(* IEC 61131-3 sources: daoli-st-library/DL_Motion (part 26) *)

(* ---- FB_DL_WindingTensionCtrl.st ---- *)
(*==============================================================================
 * 组件名称 (Component)  : FB_DL_WindingTensionCtrl
 * 所属子库 (Sublibrary) : DL_Motion
 * 当前版本 (Version)    : 1.0.1
 * 组件分类 (Category)   : 功能块（FUNCTION_BLOCK）· 卷绕工艺族 · 锥度张力闭环
 * 兼容性   (Platform)   : CODESYS 3.5 / TwinCAT 3 / 汇川 InoProShop / Schneider
 *                         Machine Expert；仅依赖 Standard.library（R_TRIG / LIMIT /
 *                         MIN / MAX / ABS / 标准类型转换）
 * 功能描述 (Function)   : 卷绕张力给定合成器。基准张力 = 目标张力 乘 锥度系数（随
 *                         机组直径由 1.0 平滑衰减到 1-K），摆辊位置误差经纯比例
 *                         修正环折算成张力修正量，两层相加后限幅输出，可直接送
 *                         比例阀或伺服转矩限幅入口。卷径可由线速度与角速度反算，
 *                         也可由外部注入。
 * 与既有件边界 (Boundary): FB_DL_WindingTraverse 做排线横动与卷径递推，不含张力
 *                         闭环；FC_DL_CoilDiameterCalc 只做单点几何反算（无状态、
 *                         无记忆）；本件是张力控制层，把二者的能力按需组装。本件
 *                         的相位枚举是工艺相位（闭环 / 开环降级），不是轴状态，轴
 *                         状态机仍归 I_DL_MotionAxis 的 PLCopen 语义，两者严禁合并。
 * 设计要点 (Key notes)  :
 *   ① 降级必须显式：摆辊反馈丢失时进 eOpenLoop 并上报 02D0，只输出锥度基准张力，
 *      不静默沿用上次闭环输出，也不静默把自己当闭环继续算；
 *   ② 修正加在基准上而非串接：摆辊失反馈时仍有锥度张力可用，失反馈不丢张力；
 *   ③ 锥度分母双重校验：满卷直径减卷芯直径小于容差即判退化，系数置 1.0 并上报
 *      01C1，绝不做出除以零的动作；系数再钳到 [1-K, 1.0]，K 自身先钳到 [0, 1]；
 *   ④ 卷径无效沿用上次有效值：转速低于门限时几何反算不可信（编码器低频量化），
 *      沿用上次有效值并累计连续无效次数，超限才升级为 02D1 锁存；
 *   ⑤ 无扰投切：开环恢复闭环时先给 PID 两拍跟踪（跟踪值 0，跟踪窗内过程值同步
 *      取基准以保偏差为零），跟踪结束积分残量为零，比例作用全量恢复；
 *      杜绝投切瞬间张力跳变；
 *   ⑥ 纯比例修正环：PID 实例积分与微分时间均给零，卷径时变工况下不会被积分饱和
 *      拖住。
 * 开源溯源 (Origin)     : 参考 lgf-technology、s7-motion 公开手册与 PLCopen 运动
 *                         控制规范中卷绕张力控制的功能分类与参数域（张力设定、锥度
 *                         系数、摆辊修正、卷径来源四段入口形态），只借分类、参数域
 *                         与命名组织，clean-room 实现，不构成衍生作品。引脚命名、
 *                         枚举、状态跃迁、故障码与合成公式 100% 自有。
 * 依赖     (Depends)    : DL_Algo 已入库件 FB_DL_PidController（拍级 PID，输出域
 *                         经 rOutMin / rOutMax 取 −1~+1 归一化）、
 *                         FC_DL_CoilDiameterCalc（几何反算，入口米制、出口米制，
 *                         本件负责毫米与米换算）。层次合法：Motion 依赖 Algo。
 * 状态迁移 (Transitions):
 *   eIdle      -- bEnable 且 bRun 且摆辊反馈有效 -----------> eClosedLoop（bInControl）
 *   eIdle      -- bEnable 且 bRun 且摆辊反馈无效 -----------> eOpenLoop（02D0 显式降级）
 *   eClosedLoop-- 摆辊反馈丢失 -----------------------------> eOpenLoop（02D0）
 *   eOpenLoop  -- 摆辊反馈连续 3 拍在物理域内 ---------------> eClosedLoop（跟踪投切）
 *   eClosedLoop-- 卷径连续无效次数超限 ---------------------> eFault（02D1 锁存）
 *   eOpenLoop  -- 卷径连续无效次数超限 ---------------------> eFault（02D1 锁存）
 *   任何运行态 -- NOT bEnable 或 NOT bRun ------------------> eIdle（输出 0，PID 复位）
 *   eFault     -- bReset 上升沿 ----------------------------> eIdle
 *   非法枚举值 -- CASE ELSE 兜底 ---------------------------> eFault（复用 02D1）
 * 码位表 (Error codes)  :
 *   16#0004_01C0【信息级】卷径无效（无有效反算或注入非法），已沿用上次有效值；
 *   16#0004_01C1【信息级】锥度系数分母退化或系数超界，已钳位；
 *   16#0004_01C2【信息级】张力输出限幅生效，输出被钳到张力域边界；
 *   16#0004_02D0【故障级】摆辊反馈丢失（非有限值或超机械行程），降级开环；
 *   16#0004_02D1【故障级】卷径连续无效超限（几何法已不可信），锁存待复位。
 *   信息级码只进 uErrorId，不置 bError；02D0 虽为故障级但只降级不停机（bError
 *   置位以提示上游），02D1 进 eFault 锁存。
 * 验收向量 (Acceptance):
 *   V1 锥度：K 0.5、卷芯 200 mm、满卷 1000 mm、实际 800 mm → 系数 0.625；
 *   V2 基准张力：同上且设定 100 N → 基准 62.5 N；
 *   V3 摆辊修正：误差 +2.0 mm、增益 0.5（归一化）、修正满量程 1.0 N → 修正 +1.0 N，
 *      输出 63.5 N；
 *   V4 满卷：实际 1000 mm、设定 100 N → 系数 0.5，基准 50.0 N；
 *   V5 卷径反算：线速 120 米每分、转速 60 转每分、直连 → 卷径约 636.6 mm；
 *   V6 卷径无效：转速 0 → 沿用上次有效卷径，码 01C0，bError 为 FALSE；
 *   V7 反馈丢失：摆辊位置 9999.0 mm → 输出等于基准（不加修正），码 02D0，
 *      bError 为 TRUE，bInControl 为 FALSE。
 * 已知限制 (Limits)     : ① 卷径反算用直连传动比 1.0（机械传动比应由卷径件入口
 *                         承载，本件不重复定义）；② 张力闭环是归一化纯比例修正，
 *                         不做卷径前馈，加减速段的动态偏差仍需现场调 fPidKp；
 *                         ③ 本件不构成安全功能，断带与超张力保护必须由硬件与
 *                         认证安全回路承担。
 * 规格偏离 (Deviation)  : ① 规格伪码把 fPidKp 原样送 PID，同时要求「摆辊正误差得
 *                         正修正」，二者符号相反；本实现送 −ABS(fPidKp)，依托 PID
 *                         件已文档化的「负增益即反作用」特性，令正误差得正修正，
 *                         与验收向量 V3 一致；② 规格成员名 nInvalidDiaCnt 定义类型
 *                         为 UDINT，与「无符号量 u 前缀」红线冲突，改名
 *                         uInvalidDiaCnt（语义不变）；③ 规格未规定故障态张力输出，
 *                         本实现取 0.0 安全值；④ 规格未覆盖「使能瞬间反馈已丢失」
 *                         路径，本实现显式进 eOpenLoop 并带 02D0，不得静默入闭环。
 * 红线自检 (Redline)    : R1 零全局变量表 / 零外部变量声明 / 零物理地址 ✓
 *                         R2 零占位符 ✓ ｜ R3 纯 IEC 61131-3 ✓
 *                         R4 防除零（锥度分母、转速门限）、防越界（卷径钳位）、
 *                         浮点容差（系数域与限幅判定）✓
 *                         R5 声明行 100% 中英双语同行注释 ✓
 *                         R6 ENUM + CASE 且 ELSE 兜底，四态各自有标签 ✓
 *                         R7 R_TRIG 与 PID 实例均在主体无条件刷新 ✓
 * 修订历史 (Revision)   :
 *   2026-11-15  v1.0.0  首版入库（Round 11 · DL_Motion 卷绕张力族开族件）
 *   2026-11-15  v1.0.1  R11 总监终审修复：跟踪拍只置位不递减（bTrack 恒真致修正恒零、
 *                       闭环退化为开环），补 eClosedLoop 逐拍递减；跟踪窗内过程值改取
 *                       基准，消除 PID 反算积分残量（原跟踪结束 fInt 恒等于负比例项，
 *                       V3 修正 +1.0 N 不可达）；02D1 判据由大于改为大于等于，与饱和
 *                       计数上限自洽（原判据在计数封顶时永假，锁存永不触发）
 *   2026-11-15  v1.0.1  R11 director final review fix: the tracking counter now decrements
 *                       every closed-loop scan, the process value follows the reference
 *                       inside the tracking window to keep the back-calculated integral at
 *                       zero, and the 02D1 test uses greater-or-equal against the
 *                       saturating counter so the latch can actually engage
 *============================================================================*)
(*-----------------------------------------------------------------------------
 * 调用示例 (Instance guide)：
 *   // fbTensionPid 与 stStat 均由调用方持有，跨周期传入
 *   fbTension(bEnable := bLineRun, bReset := bFaultReset, bRun := bWinding,
 *             fTensionSet := fTensionRecipe, fDancerPos := fDancerFeedback,
 *             fDancerRef := 0.0, fAxisSpeedRpm := fWinderRpm,
 *             fLineSpeed := fLineSpeedAct, fCoreDia := 200.0,
 *             fDiaMax := 1000.0, bUseInjectedDia := FALSE,
 *             fTaperK := 0.50, fPidKp := 0.5, fTrimSpan := 5.0,
 *             fTensionMin := 0.0, fTensionMax := 300.0);
 *   fValveCmd := fbTension.fTensionOut;
 *   注：fbTensionPid 只允许本块调用，外部不要再对该实例赋值引脚，否则归一化
 *       输出域会被覆盖，修正量会放大一百倍。
 *----------------------------------------------------------------------------*)
(*-----------------------------------------------------------------------------
 * 常见误用与现场提示 (Field notes)：
 *   1 fTaperK 给 0 表示无锥度（全程恒张力），给 1 表示满卷张力降到零，后者在
 *     实际工艺中通常不可用，建议上限取 0.7。
 *   2 摆辊反馈量程必须与 fDancerRef 同一基准：本块用绝对值 500 mm 判机械不可能
 *     值，若机械行程超过 500 mm，请把 DL_DANCER_LIMIT 调大后重新入库。
 *   3 卷径连续无效 50 次即锁存 02D1：停机不转时卷径无效属正常（信息级 01C0），
 *     只要 bRun 撤除就不会累计，现场不要把停机误判为故障。
 *   4 开环降级期间张力只随卷径变化，摆辊会漂到机械限位，现场必须给摆辊限位
 *     开关并把其信号接入上位联锁，本块不做摆辊位置保护。
 *   5 张力上下限写反时本块自动对调，但不会报警，调试期请核对 fTensionMin 与
 *     fTensionMax 的实际取值。
 *----------------------------------------------------------------------------*)
(*-----------------------------------------------------------------------------
 * 枚举: E_DL_TensionPhase（归属 DL_Motion，与本功能块同文件发布）
 * 含义: 张力工艺相位。eOpenLoop 是显式降级态而非故障态，二者不可混用。
 *----------------------------------------------------------------------------*)
{attribute 'strict'}
{attribute 'qualified_only'}
TYPE E_DL_TensionPhase :
(
    eIdle       := 0,   // 空闲：未使能或未运行，张力输出 0，PID 复位 / Idle: disabled or not running, tension output zero, PID reset
    eOpenLoop   := 10,  // 开环降级：摆辊反馈不可用，只出锥度基准张力 / Open loop degraded: dancer feedback unusable, taper base only
    eClosedLoop := 20,  // 闭环运行：基准张力加摆辊比例修正 / Closed loop: base tension plus dancer proportional trim
    eFault      := 99   // 故障锁存：卷径几何法不可信，仅复位沿退出 / Fault latched: diameter geometry untrusted, exits on reset edge only
) UINT;
END_TYPE
(*-----------------------------------------------------------------------------
 * 结构体: ST_DL_WindingStat（归属 DL_Motion，与本功能块同文件发布）
 * 含义: 卷绕统计，由调用方持有并可持久化到配方域。
 *----------------------------------------------------------------------------*)
TYPE ST_DL_WindingStat :
STRUCT
    fTensionAvg     : REAL;   // 张力滑动均值 [N]，一阶指数平均，仅闭环期更新 / Tension running average in newtons, updated in closed loop only
    uInvalidDiaCnt  : UDINT;  // 卷径连续无效次数 [次]，任一有效反算即清零 / Consecutive invalid diameter count, cleared by any valid result
    tRunTime        : TIME;   // 闭环累计运行时长 [ms]，按任务周期累加 / Accumulated closed-loop runtime in milliseconds
END_STRUCT
END_TYPE

(*==============================================================================
 * 功能块: FB_DL_WindingTensionCtrl
 * 调用约定: 每扫描周期无条件调用一次；PID 实例在主体末尾无条件调用。
 * 无状态泄漏: 状态驻留实例私有 VAR 与调用方持有的 stStat / fbTensionPid。
 *============================================================================*)
FUNCTION_BLOCK FB_DL_WindingTensionCtrl
VAR_INPUT
    bEnable          : BOOL := FALSE;        // 总使能 [BOOL]，FALSE 时输出 0 并复位 PID / Master enable, FALSE zeroes the output and resets the PID
    bReset           : BOOL := FALSE;        // 复位 [BOOL]，上升沿复位故障、计数与 PID / Reset, rising edge clears fault, counters and the PID
    bRun             : BOOL := FALSE;        // 卷绕运行中 [BOOL]，FALSE 时张力给定保持 0 / Winding running flag, FALSE holds the tension command at zero
    fTensionSet      : REAL := 0.0;          // 目标张力（满卷前基准）[N]，域 0.0~500.0 / Base tension setpoint in newtons, range zero to five hundred
    fDancerPos       : REAL := 0.0;          // 摆辊实际位置 [mm]，0 为机械中位，绝对值超 500 判失效 / Dancer actual position in millimetres, zero at mechanical centre
    fDancerRef       : REAL := 0.0;          // 摆辊中位基准 [mm]，非有限值按 0 处理 / Dancer centre reference in millimetres, non-finite treated as zero
    fAxisSpeedRpm    : REAL := 0.0;          // 卷轴转速 [转每分]，低于 1.0 视为不可反算 / Winder shaft speed in revolutions per minute, below one is untrusted
    fLineSpeed       : REAL := 0.0;          // 线速度 [米每分]，与卷径件入口同单位 / Line speed in metres per minute, same unit as the diameter function input
    fCoreDia         : REAL := 200.0;        // 卷芯直径 [mm]，域 10.0~3000.0 / Core diameter in millimetres, range ten to three thousand
    fDiaMax          : REAL := 1000.0;       // 满卷直径 [mm]，必须大于卷芯直径，否则锥度退化 / Full roll diameter in millimetres, must exceed the core diameter
    fDiaInjected     : REAL := 0.0;          // 外部注入卷径 [mm]，视觉或上位机来源 / Injected diameter in millimetres from vision or a host system
    bUseInjectedDia  : BOOL := FALSE;        // 卷径来源选择 [BOOL]，TRUE 用注入值，FALSE 由速度比反算 / Diameter source, TRUE uses the injected value
    fThickness       : REAL := 0.10;         // 材料厚度 [mm]，供卷径件层数积分 / Material thickness in millimetres, used by the layer integral
    fTaperK          : REAL := 0.50;         // 锥度系数 [无量纲 0~1]，满卷张力降至 1-K 倍 / Taper coefficient, full roll tension falls to one minus K
    fPidKp           : REAL := 0.5;          // 摆辊修正归一化增益 [每毫米]，输出域 −1~+1，取绝对值后反作用 / Normalised dancer gain per millimetre, absolute value used with reverse action
    fTrimSpan        : REAL := 1.0;          // 修正满量程 [N]，归一化输出乘该值即张力修正 / Trim span in newtons, the normalised output multiplied by this value
    fTensionMin      : REAL := 0.0;          // 张力输出下限 [N]，与上限对调时自动修复 / Tension lower limit in newtons, swapped limits are repaired
    fTensionMax      : REAL := 500.0;        // 张力输出上限 [N]，等于下限时输出被钉死 / Tension upper limit in newtons, an equal limit pins the output
END_VAR
VAR_OUTPUT
    fTensionOut      : REAL := 0.0;          // 张力给定输出 [N]，送比例阀或转矩限幅入口 / Tension command output in newtons for a proportional valve or torque limit
    fDiaAct          : REAL := 0.0;          // 当前生效卷径 [mm]，已钳入物理域 / Effective diameter in millimetres, clamped into the physical range
    fTaperFactor     : REAL := 1.0;          // 实际锥度系数 [无量纲]，域 1-K~1.0 / Effective taper factor, range one minus K to one
    fDancerErr       : REAL := 0.0;          // 摆辊位置误差 [mm]，等于实测减基准 / Dancer position error in millimetres, measured minus reference
    eState           : E_DL_TensionPhase := E_DL_TensionPhase.eIdle; // 主状态机当前态 [枚举] / Current state of the main state machine
    bInControl       : BOOL := FALSE;        // 张力闭环生效 [BOOL]，仅 eClosedLoop 为 TRUE / Closed-loop tension active, TRUE only in the closed-loop state
    bError           : BOOL := FALSE;        // 故障标志 [BOOL]，故障级码或降级态置位，信息级码不置位 / Fault flag, set by fault-level codes or the degraded state
    uErrorId         : UDINT := 0;           // 事件或故障码 [段位 0004_01Cx 与 0004_02Dx]，0 表示无事件 / Event or fault code in the 0004 bands, zero means none
    fDiaLastValid    : REAL := 0.0;          // 最近一次有效卷径 [mm]，0 表示尚无有效值 / Last valid diameter in millimetres, zero means none yet
END_VAR
VAR_IN_OUT
    fbTensionPid     : FB_DL_PidController;  // 摆辊修正环 PID 实例 [FB]，由调用方持有且只允许本块调用 / Dancer trim PID instance held by the caller and driven only by this block
    stStat           : ST_DL_WindingStat;    // 跨周期卷绕统计 [结构体]，由调用方持有 / Persistent winding statistics held by the caller
END_VAR
VAR
    bInit            : BOOL := FALSE;        // 首扫完成标志 [BOOL]，初值 FALSE，判据恒为 NOT bInit / First-scan done flag, initial FALSE, judged by NOT bInit
    bDancerOk        : BOOL := FALSE;        // 摆辊反馈有效判据 [BOOL]，逐拍重算 / Dancer feedback verdict, recomputed every scan
    bDancerLost      : BOOL := FALSE;        // 摆辊反馈丢失标志 [BOOL]，降级原因量 / Dancer feedback lost flag, the explicit degradation reason
    bAvgInit         : BOOL := FALSE;        // 张力均值首样本标志 [BOOL]，避免从 0 起算 / Tension average first-sample flag, avoids averaging from zero
    nRecoverCnt      : INT := 0;             // 反馈恢复连续拍计数 [拍]，满 3 拍回闭环 / Consecutive good-feedback counter, three scans restore closed loop
    nTrackSync       : INT := 0;             // 投切跟踪剩余拍数 [拍]，大于 0 时 PID 跟踪 / Remaining tracking scans, the PID tracks while above zero
    fDancerPosEff    : REAL := 0.0;          // 喂给 PID 的摆辊位置 [mm]，失效时以基准值替代 / Dancer position fed to the PID, replaced by the reference when invalid
    fDancerRefEff    : REAL := 0.0;          // 生效摆辊基准 [mm]，已做非有限值防御 / Effective dancer reference after the non-finite defence
    fPidPvEff        : REAL := 0.0;          // 喂给 PID 的过程值 [mm]，跟踪窗口内以基准替代 / Process value fed to the PID, replaced by the reference inside the tracking window
    fTensionSetEff   : REAL := 0.0;          // 生效目标张力 [N]，已做非有限值防御 / Effective tension setpoint after the non-finite defence
    fTrimSpanEff     : REAL := 1.0;          // 生效修正满量程 [N]，取绝对值 / Effective trim span in newtons, absolute value used
    fPidKpEff        : REAL := 0.0;          // 送入 PID 的增益 [每毫米]，取负值实现反作用 / Gain passed to the PID, negated for reverse action
    fCoreDiaEff      : REAL := 200.0;        // 生效卷芯直径 [mm]，钳入物理域 / Effective core diameter in millimetres, clamped into the physical range
    fDiaMaxEff       : REAL := 1000.0;       // 生效满卷直径 [mm]，钳入物理域 / Effective full-roll diameter in millimetres, clamped into the physical range
    fTaperKEff       : REAL := 0.50;         // 生效锥度系数 [无量纲 0~1]，越界钳位 / Effective taper coefficient, clamped into zero to one
    fTaperLow        : REAL := 0.50;         // 锥度系数下限 [无量纲]，等于 1 减生效锥度 / Taper factor lower bound, equal to one minus the effective coefficient
    fTaperRaw        : REAL := 1.0;          // 未钳位的锥度系数 [无量纲]，用于超界判定 / Unclamped taper factor used for the out-of-range test
    fDiaCalc         : REAL := 0.0;          // 卷径反算结果 [mm]，已做米转毫米 / Diameter result in millimetres after the metre conversion
    fDiaLReal        : LREAL := 0.0;         // 卷径件出口绑定值 [米]，LREAL 精度承接 / Diameter bound from the function output in metres at LREAL precision
    fDiaRet          : LREAL := 0.0;         // 卷径件返回值 [米]，函数返回即滤波后卷径 / Diameter function return value in metres, the filtered diameter
    fBase            : REAL := 0.0;          // 锥度基准张力 [N]，等于设定乘锥度系数 / Taper base tension in newtons, setpoint times the taper factor
    fTrim            : REAL := 0.0;          // 摆辊张力修正 [N]，闭环时等于归一化输出乘满量程 / Dancer trim in newtons, the normalised output times the span
    fRawCmd          : REAL := 0.0;           // 未限幅的张力指令 [N]，限幅前中间量 / Unlimited tension command in newtons before clamping
    fLimLow          : REAL := 0.0;          // 生效张力下限 [N]，已做上下对调修复 / Effective tension lower limit after repair
    fLimHigh         : REAL := 500.0;        // 生效张力上限 [N]，已做上下对调修复 / Effective tension upper limit after repair
    fAvgAlpha        : REAL := 0.0;          // 张力均值一阶权重 [无量纲]，由任务周期与时间常数算出 / First-order weight of the tension average
    uErrInfo         : UDINT := 0;           // 本拍瞬时信息码 [段位 0004_01C0~01C2]，逐拍重算 / Transient info code recomputed every scan
    uErrFault        : UDINT := 0;           // 锁存故障码 [段位 0004_02D1]，仅复位清除 / Latched fault code, cleared by reset only
    fbTrigReset      : R_TRIG;               // 复位上升沿检测实例 / Rising edge detector for the reset flag
    fbTrigRun        : R_TRIG;               // 运行上升沿检测实例 / Rising edge detector for the running flag
END_VAR
VAR CONSTANT
    DL_FLOAT_EPS     : REAL := 1.0E-6;       // 浮点判等与判零容差 [无量纲，按比较量量纲同值使用] / Float equality and zero tolerance
    DL_INF_MAX       : REAL := 1.0E30;       // 有限值幅值上限 [无量纲，按各量量纲同值使用] / Finite magnitude upper bound
    DL_RPM_MIN       : REAL := 1.0;          // 卷径反算最小转速 [转每分]，低于此值不反算 / Minimum speed for the inverse diameter calculation
    DL_DIA_MIN       : REAL := 10.0;         // 卷径物理下限 [mm] / Diameter physical lower bound in millimetres
    DL_DIA_MAX       : REAL := 3000.0;       // 卷径物理上限 [mm] / Diameter physical upper bound in millimetres
    DL_DANCER_LIMIT  : REAL := 500.0;        // 摆辊机械行程上限 [mm]，绝对值超此判失效 / Dancer mechanical travel bound in millimetres
    DL_TASK_CYCLE    : REAL := 0.010;        // 主任务周期 [s]，供卷径件变化率换算 / Main task cycle in seconds for the diameter rate
    DL_TASK_TIME     : TIME := T#10MS;       // 主任务周期时间量 [ms]，供运行时长累加 / Main task cycle as a time value for runtime accumulation
    DL_FILTER_TAU    : REAL := 0.50;         // 卷径一阶低通时间常数 [s] / Diameter low-pass time constant in seconds
    DL_INVALID_MAX   : UDINT := 50;          // 卷径连续无效次数上限 [次]，超限锁存 02D1 / Consecutive invalid diameter limit before latching
    DL_RECOVER_N     : INT := 3;             // 反馈恢复确认拍数 [拍]，连续满足才回闭环 / Consecutive good scans required to restore the closed loop
    DL_AVG_TAU       : REAL := 1.0;          // 张力均值时间常数 [s]，一阶平均用 / Tension average time constant in seconds
END_VAR
(*------------------------------------------------------------------------------
 * 段 1｜边沿实例无条件周期刷新（红线 R7：严禁置于 IF 或 CASE 分支内）｜Unconditional edge refresh, never placed inside IF or CASE branches
 *-----------------------------------------------------------------------------*)
fbTrigReset(CLK := bReset);
fbTrigRun(CLK := bRun);
(*------------------------------------------------------------------------------
 * 段 2｜瞬时输出与瞬时码预清零（出口只置位，跨拍残留一律在入口清）｜Pre-clear transient outputs and info codes at scan entry
 *-----------------------------------------------------------------------------*)
bInControl := FALSE;                        // 闭环生效标志预清零 [BOOL] / Pre-clear the closed-loop flag
fTrim      := 0.0;                          // 修正量预清零，开环与空闲不得继承上次值 [N] / Pre-clear the trim so open loop never inherits it
uErrInfo   := 0;                            // 瞬时信息码预清零 [码] / Pre-clear the transient info code
(*------------------------------------------------------------------------------
 * 段 3｜参数域修复（引脚可在线改，故逐拍重算；域非法只钳位不锁存）｜Parameter domain repair, clamping only without latching
 *-----------------------------------------------------------------------------*)
IF fTensionMax < fTensionMin THEN
    fLimLow  := fTensionMax;                // 张力域上下对调修复：下限取原上限 [N] / Repaired lower limit takes the original upper
    fLimHigh := fTensionMin;                // 张力域上下对调修复：上限取原下限 [N] / Repaired upper limit takes the original lower
ELSE
    fLimLow  := fTensionMin;                // 合法下限直通 [N] / Valid lower limit passed through
    fLimHigh := fTensionMax;                // 合法上限直通 [N] / Valid upper limit passed through
END_IF

IF (fTensionSet <> fTensionSet) OR (ABS(fTensionSet) > DL_INF_MAX) THEN
    fTensionSetEff := 0.0;                  // 目标张力非有限 → 0，宁可失张力也不给非法值 [N] / Non-finite setpoint falls back to zero
ELSE
    fTensionSetEff := fTensionSet;          // 合法目标张力直通 [N] / Valid setpoint passed through
END_IF

IF (fTrimSpan <> fTrimSpan) OR (ABS(fTrimSpan) > DL_INF_MAX) THEN
    fTrimSpanEff := 0.0;                    // 修正满量程非有限 → 0，等效关闭摆辊修正 [N] / Non-finite trim span disables the dancer trim
ELSE
    fTrimSpanEff := ABS(fTrimSpan);         // 修正满量程取绝对值 [N] / Absolute trim span
END_IF
// 送入 PID 的增益取负实现反作用：摆辊正误差（上偏）对应增张力，与验收向量 V3 一致
IF (fPidKp <> fPidKp) OR (ABS(fPidKp) > DL_INF_MAX) THEN
    fPidKpEff := 0.0;                       // 增益非有限 → 0，等效关闭修正 [每毫米] / Non-finite gain disables the trim
ELSE
    fPidKpEff := -ABS(fPidKp);              // 取绝对值后取负，负增益即 PID 件的反作用语义 [每毫米] / Absolute value negated for reverse action
END_IF

IF (fDancerRef <> fDancerRef) OR (ABS(fDancerRef) > DL_DANCER_LIMIT) THEN
    fDancerRefEff := 0.0;                   // 摆辊基准非法 → 回机械中位 0 [mm] / Illegal reference falls back to the mechanical centre
ELSE
    fDancerRefEff := fDancerRef;            // 合法基准直通 [mm] / Valid reference passed through
END_IF

IF (fCoreDia <> fCoreDia) OR (ABS(fCoreDia) > DL_INF_MAX) THEN
    fCoreDiaEff := DL_DIA_MIN;              // 卷芯直径非法 → 回物理下限 [mm] / Illegal core diameter falls back to the physical lower bound
ELSE
    fCoreDiaEff := LIMIT(DL_DIA_MIN, fCoreDia, DL_DIA_MAX); // 卷芯直径钳入物理域 [mm] / Core diameter clamped into the physical range
END_IF

IF (fDiaMax <> fDiaMax) OR (ABS(fDiaMax) > DL_INF_MAX) THEN
    fDiaMaxEff := DL_DIA_MAX;               // 满卷直径非法 → 回物理上限 [mm] / Illegal full-roll diameter falls back to the physical upper bound
ELSE
    fDiaMaxEff := LIMIT(DL_DIA_MIN, fDiaMax, DL_DIA_MAX);   // 满卷直径钳入物理域 [mm] / Full-roll diameter clamped into the physical range
END_IF
// 锥度系数域校验：非有限或越出 0~1 一律钳位并置信息级 01C1，绝不带非法系数进公式
IF (fTaperK <> fTaperK) OR (ABS(fTaperK) > DL_INF_MAX) THEN
    fTaperKEff := 0.0;                      // 非有限系数按无锥度处理，先判非数再钳位，避免 NaN 穿过 LIMIT [无量纲] / Non-finite coefficient treated as no taper
    IF bEnable AND bRun THEN
        uErrInfo := 16#0004_01C1;           // 【信息级】锥度系数非有限已按无锥度处理 / Info: non-finite taper coefficient replaced
    END_IF
ELSIF (fTaperK < 0.0) OR (fTaperK > 1.0) THEN
    fTaperKEff := LIMIT(0.0, fTaperK, 1.0); // 越界钳到 0~1 双向钳位 [无量纲] / Two-sided clamp into zero to one
    IF bEnable AND bRun THEN
        uErrInfo := 16#0004_01C1;           // 【信息级】锥度系数超界已钳位 / Info: taper coefficient clamped
    END_IF
ELSE
    fTaperKEff := fTaperK;                  // 合法锥度系数直通 [无量纲] / Valid taper coefficient passed through
END_IF
// 张力均值一阶权重：由任务周期与时间常数算出，分母恒正（时间常数有下限保证）
fAvgAlpha := DL_TASK_CYCLE / (DL_AVG_TAU + DL_TASK_CYCLE); // 均值权重 [无量纲] / First-order average weight
(*------------------------------------------------------------------------------
 * 段 4｜首扫装载（R19 唯一合法范式：bInit 初值 FALSE，判据 NOT bInit）｜First-scan load, the only accepted initialisation pattern
 *-----------------------------------------------------------------------------*)
IF NOT bInit THEN
    stStat.fTensionAvg    := 0.0;           // 张力均值清零，等首个闭环样本直取 [N] / Clear the tension average until the first closed-loop sample
    stStat.uInvalidDiaCnt := 0;             // 卷径无效计数清零 [次] / Clear the invalid diameter counter
    stStat.tRunTime       := T#0S;          // 运行时长清零 [ms] / Clear the accumulated runtime
    fDiaLastValid         := 0.0;           // 有效卷径历史清零，0 表示尚无有效值 [mm] / Clear the valid diameter history
    bDancerLost           := FALSE;         // 反馈丢失标志清零 [BOOL] / Clear the feedback lost flag
    nRecoverCnt           := 0;             // 恢复计数清零 [拍] / Clear the recovery counter
    nTrackSync            := 0;             // 投切跟踪计数清零 [拍] / Clear the tracking counter
    bAvgInit              := FALSE;         // 均值首样本标志清零 [BOOL] / Clear the average first-sample flag
    bInit                 := TRUE;          // 首扫完成置位 [BOOL] / First scan completed
END_IF
(*------------------------------------------------------------------------------
 * 段 5｜复位（清故障、计数与降级标志；PID 由复位引脚同步清除；参数域不动）｜Reset clears the latched fault, counters and degradation flags
 *-----------------------------------------------------------------------------*)
IF fbTrigReset.Q THEN
    uErrFault             := 0;             // 锁存故障码清零 [码] / Clear the latched fault code
    uErrInfo              := 0;             // 瞬时信息码清零 [码] / Clear the transient info code
    stStat.uInvalidDiaCnt := 0;             // 卷径无效计数清零，允许重新起步 [次] / Clear the invalid diameter counter so production can restart
    bDancerLost           := FALSE;         // 反馈丢失标志清零 [BOOL] / Clear the feedback lost flag
    nRecoverCnt           := 0;             // 恢复计数清零 [拍] / Clear the recovery counter
    nTrackSync            := 0;             // 跟踪计数清零 [拍] / Clear the tracking counter
    eState                := E_DL_TensionPhase.eIdle; // 回空闲，等待使能与运行条件 [枚举] / Back to idle waiting for enable and run
END_IF

IF fbTrigRun.Q THEN
    bAvgInit := FALSE;                      // 新一次卷绕启动：张力均值重新直取首样本，不继承上一卷 [BOOL] / New run restarts the tension average instead of inheriting the last roll
END_IF
(*------------------------------------------------------------------------------
 * 段 6｜摆辊反馈有效性判定（非有限值或超机械行程即判失效，显式标记原因）｜Dancer feedback verdict with an explicit reason flag
 *-----------------------------------------------------------------------------*)
bDancerOk := NOT ((fDancerPos <> fDancerPos) OR (ABS(fDancerPos) > DL_DANCER_LIMIT));
IF bDancerOk THEN
    fDancerPosEff := fDancerPos;            // 有效反馈直通，喂给 PID [mm] / Valid feedback passed through to the PID
ELSE
    fDancerPosEff := fDancerRefEff;         // 失效反馈以基准替代，令 PID 偏差为零且 NaN 不扩散 [mm] / Substitute the reference so the PID error stays zero
END_IF
fDancerErr := fDancerPosEff - fDancerRefEff; // 摆辊位置误差，实测减基准 [mm] / Dancer position error, measured minus reference
(*------------------------------------------------------------------------------
 * 段 7｜卷径获取（注入优先；否则按速度比反算；无效沿用上次有效值并计数）｜Diameter acquisition with reuse-on-invalid and consecutive counting
 *-----------------------------------------------------------------------------*)
IF bEnable AND bRun THEN
    IF bUseInjectedDia THEN
        IF (fDiaInjected <> fDiaInjected) OR (ABS(fDiaInjected) > DL_INF_MAX) THEN
            IF fDiaLastValid > DL_FLOAT_EPS THEN
                fDiaAct := fDiaLastValid;   // 注入值非法 → 沿用上次有效卷径 [mm] / Illegal injection reuses the last valid diameter
            ELSE
                fDiaAct := fCoreDiaEff;     // 无历史有效值 → 以卷芯直径兜底，杜绝零卷径除零 [mm] / Fall back to the core diameter when no history exists
            END_IF
            IF stStat.uInvalidDiaCnt < DL_INVALID_MAX THEN
                stStat.uInvalidDiaCnt := stStat.uInvalidDiaCnt + 1; // 连续无效计数累加，封顶后靠 02D1 锁存 [次] / Saturating invalid counter
            END_IF
            uErrInfo := 16#0004_01C0;       // 【信息级】卷径无效已沿用上次有效值 / Info: invalid diameter, last valid value reused
        ELSE
            fDiaAct := LIMIT(DL_DIA_MIN, fDiaInjected, DL_DIA_MAX); // 注入卷径钳入物理域 [mm] / Injected diameter clamped into the physical range
            IF (fDiaInjected < DL_DIA_MIN) OR (fDiaInjected > DL_DIA_MAX) THEN
                uErrInfo := 16#0004_01C0;   // 【信息级】注入卷径超物理域已钳位 / Info: injected diameter clamped
            END_IF
            fDiaLastValid         := fDiaAct; // 记录有效卷径 [mm] / Record the valid diameter
            stStat.uInvalidDiaCnt := 0;     // 有效值出现即清零连续无效计数 [次] / Reset the consecutive counter on any valid value
        END_IF
    ELSE
        IF (fAxisSpeedRpm <> fAxisSpeedRpm) OR (ABS(fAxisSpeedRpm) > DL_INF_MAX)
           OR (fAxisSpeedRpm < DL_RPM_MIN)
           OR (fLineSpeed <> fLineSpeed) OR (ABS(fLineSpeed) > DL_INF_MAX) THEN
            IF fDiaLastValid > DL_FLOAT_EPS THEN
                fDiaAct := fDiaLastValid;   // 低速或入参非法 → 沿用上次有效卷径 [mm] / Low speed or illegal input reuses the last valid diameter
            ELSE
                fDiaAct := fCoreDiaEff;     // 无历史有效值 → 以卷芯直径兜底 [mm] / Fall back to the core diameter
            END_IF
            IF stStat.uInvalidDiaCnt < DL_INVALID_MAX THEN
                stStat.uInvalidDiaCnt := stStat.uInvalidDiaCnt + 1; // 连续无效计数累加 [次] / Saturating invalid counter
            END_IF
            uErrInfo := 16#0004_01C0;       // 【信息级】卷径无效已沿用上次有效值 / Info: invalid diameter, last valid value reused
        ELSE
            // 按已入库卷径件的真实契约调用：入口为米制与秒制，出口绑定滤波后卷径（米）
            fDiaRet := FC_DL_CoilDiameterCalc(
                fLineSpeed := REAL_TO_LREAL(fLineSpeed),              // 米每分，与本件引脚同单位 / Metres per minute, same unit as this pin
                fShaftRpm  := REAL_TO_LREAL(fAxisSpeedRpm),           // 转每分，与卷轴转速同单位 / Revolutions per minute
                fGearRatio := 1.0,                                    // 直连，机械传动比由卷径件入口承载 / Direct drive, the gear ratio belongs to the function input
                fCoreDia   := REAL_TO_LREAL(fCoreDiaEff) / 1000.0,     // 毫米转米 / Millimetres converted to metres
                fThickness := REAL_TO_LREAL(fThickness) / 1000.0,     // 毫米转米 / Millimetres converted to metres
                fPrevDia   := REAL_TO_LREAL(fDiaLastValid) / 1000.0,  // 毫米转米，0 表示无历史 / Millimetres converted to metres, zero means no history
                fTaskCycle := REAL_TO_LREAL(DL_TASK_CYCLE),           // 任务周期，秒 / Task cycle in seconds
                bFilterEn  := TRUE,                                   // 卷径低通使能 / Diameter low-pass enabled
                fFilterTau := REAL_TO_LREAL(DL_FILTER_TAU),           // 低通时间常数，秒 / Low-pass time constant in seconds
                fDia       => fDiaLReal );                            // 出口绑定：滤波后卷径，米 / Bound output, filtered diameter in metres
            fDiaCalc := LREAL_TO_REAL(fDiaLReal * 1000.0);            // 米转毫米，显式转换，出口绑定优先 / Metres converted to millimetres, the bound output is preferred
            IF (fDiaLReal <> fDiaLReal) AND (fDiaRet = fDiaRet) THEN
                fDiaCalc := LREAL_TO_REAL(fDiaRet * 1000.0);          // 绑定值非法而返回值有效 → 退回返回值，兼容平台绑定差异 / Bound value illegal, fall back to the function return
            END_IF
            IF (fDiaCalc <> fDiaCalc) OR (fDiaCalc <= DL_FLOAT_EPS) THEN
                IF fDiaLastValid > DL_FLOAT_EPS THEN
                    fDiaAct := fDiaLastValid; // 反算结果不可用 → 沿用上次有效卷径 [mm] / Unusable result reuses the last valid diameter
                ELSE
                    fDiaAct := fCoreDiaEff;   // 无历史有效值 → 以卷芯直径兜底 [mm] / Fall back to the core diameter
                END_IF
                IF stStat.uInvalidDiaCnt < DL_INVALID_MAX THEN
                    stStat.uInvalidDiaCnt := stStat.uInvalidDiaCnt + 1; // 连续无效计数累加 [次] / Saturating invalid counter
                END_IF
                uErrInfo := 16#0004_01C0;   // 【信息级】反算结果不可用已沿用上次有效值 / Info: unusable result, last valid value reused
            ELSE
                fDiaAct := LIMIT(DL_DIA_MIN, fDiaCalc, DL_DIA_MAX); // 反算卷径钳入物理域 [mm] / Computed diameter clamped into the physical range
                fDiaLastValid         := fDiaAct; // 记录有效卷径 [mm] / Record the valid diameter
                stStat.uInvalidDiaCnt := 0;       // 有效反算即清零连续无效计数 [次] / Reset the consecutive counter on a valid result
            END_IF
        END_IF
    END_IF
ELSE
    IF fDiaLastValid > DL_FLOAT_EPS THEN
        fDiaAct := fDiaLastValid;           // 非运行态不反算，沿用上次有效卷径 [mm] / Not running, reuse the last valid diameter
    ELSE
        fDiaAct := fCoreDiaEff;             // 非运行且无历史 → 以卷芯直径兜底 [mm] / Not running without history falls back to the core diameter
    END_IF
END_IF

// 卷径输出钳位兜底：任何路径都不得把非法值送出（防御性二次确认）
IF (fDiaAct <> fDiaAct) OR (fDiaAct < DL_DIA_MIN) OR (fDiaAct > DL_DIA_MAX) THEN
    fDiaAct := LIMIT(DL_DIA_MIN, fDiaAct, DL_DIA_MAX); // 卷径域二次钳位 [mm] / Second-stage diameter clamp
    IF fDiaAct <> fDiaAct THEN
        fDiaAct := fCoreDiaEff;             // 仍为非法值 → 回卷芯直径 [mm] / Still illegal, fall back to the core diameter
    END_IF
END_IF
(*------------------------------------------------------------------------------
 * 段 8｜锥度系数（分母双重校验，系数双向钳位，退化或超界置 01C1）｜Taper factor with denominator guard and two-sided clamping
 *-----------------------------------------------------------------------------*)
IF ABS(fDiaMaxEff - fCoreDiaEff) <= DL_FLOAT_EPS THEN
    fTaperFactor := 1.0;                    // 满卷等于卷芯：锥度退化，系数取 1.0 防除零 [无量纲] / Degenerate span, unity factor avoids division by zero
    IF bEnable AND bRun THEN
        uErrInfo := 16#0004_01C1;           // 【信息级】锥度分母退化已改置 1.0 / Info: degenerate taper span replaced by unity
    END_IF
ELSE
    fTaperLow := 1.0 - fTaperKEff;          // 锥度系数下限，等于 1 减锥度 [无量纲] / Taper factor lower bound
    fTaperRaw := 1.0 - fTaperKEff * (fDiaAct - fCoreDiaEff) / (fDiaMaxEff - fCoreDiaEff); // 原始锥度系数 [无量纲] / Raw taper factor
    IF (fTaperRaw > 1.0 + DL_FLOAT_EPS) OR (fTaperRaw < fTaperLow - DL_FLOAT_EPS) THEN
        fTaperFactor := LIMIT(fTaperLow, fTaperRaw, 1.0); // 超界钳到 [1-K, 1] [无量纲] / Clamp into the lower bound and one
        IF bEnable AND bRun THEN
            uErrInfo := 16#0004_01C1;       // 【信息级】锥度系数超界已钳位 / Info: taper factor clamped
        END_IF
    ELSE
        fTaperFactor := fTaperRaw;          // 未超界直通 [无量纲] / Raw factor passed through
    END_IF
END_IF
(*------------------------------------------------------------------------------
 * 段 9｜锥度基准张力（修正项后续加在基准上，失反馈也不丢张力）｜Taper base tension, the trim is added on top later
 *-----------------------------------------------------------------------------*)
fBase := fTensionSetEff * fTaperFactor;     // 基准张力＝目标张力乘锥度系数 [N] / Base tension equals setpoint times taper factor
(*------------------------------------------------------------------------------
 * 段 10｜主状态机（红线 R6：ENUM + CASE + ELSE 兜底，四态各有标签）｜Main state machine with mandatory ELSE fallback and four labelled states
 *-----------------------------------------------------------------------------*)
CASE eState OF

    E_DL_TensionPhase.eIdle:                // 空闲：等使能与运行条件，张力输出在段 12 强制为 0
        IF bEnable AND bRun THEN
            IF bDancerOk THEN
                nTrackSync  := 2;           // 无扰投切：先给 PID 两拍跟踪 [拍] / Two tracking scans for a bumpless transfer
                bDancerLost := FALSE;       // 反馈有效，降级原因清除 [BOOL] / Feedback valid, clear the degradation reason
                eState      := E_DL_TensionPhase.eClosedLoop;
            ELSE
                bDancerLost := TRUE;        // 显式记录降级原因：反馈缺失 [BOOL] / Record the explicit degradation reason
                nRecoverCnt := 0;           // 恢复计数从零开始 [拍] / Recovery counter starts at zero
                eState      := E_DL_TensionPhase.eOpenLoop; // 使能瞬间反馈已失效，直接进降级态 [枚举] / Enter the degraded state directly
            END_IF
        END_IF

    E_DL_TensionPhase.eClosedLoop:          // 闭环运行：基准加摆辊比例修正
        IF nTrackSync > 0 THEN
            nTrackSync := nTrackSync - 1;   // 跟踪拍递减，减到零才放开修正 [拍] / Decrement the tracking counter until the trim is released
        END_IF
        IF (NOT bEnable) OR (NOT bRun) THEN
            nTrackSync := 0;                // 停机撤跟踪 [拍] / Clear the tracking counter on stop
            eState     := E_DL_TensionPhase.eIdle;
        ELSIF stStat.uInvalidDiaCnt >= DL_INVALID_MAX THEN
            uErrFault := 16#0004_02D1;      // 【故障级】卷径连续无效超限，几何法不可信 / Fault: consecutive invalid diameters exceeded the limit
            eState    := E_DL_TensionPhase.eFault;
        ELSIF NOT bDancerOk THEN
            bDancerLost := TRUE;            // 显式降级：反馈丢失 [BOOL] / Explicit degradation on feedback loss
            nRecoverCnt := 0;               // 恢复计数重新开始 [拍] / Recovery counter restarts
            nTrackSync  := 0;               // 撤闭环跟踪 [拍] / Clear the closed-loop tracking counter
            eState      := E_DL_TensionPhase.eOpenLoop;
        END_IF

    E_DL_TensionPhase.eOpenLoop:            // 开环降级：只出锥度基准张力，修正恒为 0
        IF (NOT bEnable) OR (NOT bRun) THEN
            bDancerLost := FALSE;           // 停机清降级原因 [BOOL] / Clear the degradation reason on stop
            nRecoverCnt := 0;               // 恢复计数清零 [拍] / Clear the recovery counter
            eState      := E_DL_TensionPhase.eIdle;
        ELSIF stStat.uInvalidDiaCnt >= DL_INVALID_MAX THEN
            uErrFault := 16#0004_02D1;      // 【故障级】卷径连续无效超限 / Fault: consecutive invalid diameters exceeded the limit
            eState    := E_DL_TensionPhase.eFault;
        ELSIF bDancerOk THEN
            nRecoverCnt := nRecoverCnt + 1; // 连续有效拍数累加 [拍] / Count the consecutive good scans
            IF nRecoverCnt >= DL_RECOVER_N THEN
                nRecoverCnt := 0;           // 恢复确认后计数归零 [拍] / Reset the counter after confirmation
                nTrackSync  := 2;           // 回闭环先跟踪两拍，修正从 0 起爬 [拍] / Track for two scans so the trim starts from zero
                bDancerLost := FALSE;       // 降级原因清除 [BOOL] / Clear the degradation reason
                eState      := E_DL_TensionPhase.eClosedLoop;
            END_IF
        ELSE
            nRecoverCnt := 0;               // 反馈再次失效，恢复计数归零 [拍] / Feedback failed again, reset the counter
        END_IF

    E_DL_TensionPhase.eFault:               // 故障锁存：输出安全值，仅复位沿退出
        bInControl := FALSE;                // 故障态闭环必然未生效 [BOOL] / Closed loop is not active in the fault state
        fTrim      := 0.0;                  // 故障态修正清零 [N] / Clear the trim in the fault state

    ELSE                                    // 非法状态兜底：复用本件最高优先故障码，不另造码
        uErrFault  := 16#0004_02D1;         // 【故障级】非法状态兜底，复用 02D1 / Fault: illegal state fallback reusing 02D1
        eState     := E_DL_TensionPhase.eFault;
        bInControl := FALSE;                // 强制非闭环 [BOOL] / Force the loop inactive
        fTrim      := 0.0;                  // 修正清零 [N] / Clear the trim

END_CASE
(*------------------------------------------------------------------------------
 * 段 11｜摆辊修正环实例无条件调用（FB 实例严禁放在 IF 或 CASE 分支内）｜Unconditional PID call, normalised output, pure proportional action
 *-----------------------------------------------------------------------------*)
// 跟踪窗口内以基准替代过程值：偏差恒为零，PID 反算积分保持零，窗口结束即恢复全量比例作用
// Inside the tracking window the reference replaces the process value: the error stays zero,
// so the back-calculated integral stays zero and full proportional action resumes afterwards
fPidPvEff := fDancerPosEff;
IF nTrackSync > 0 THEN
    fPidPvEff := fDancerRefEff;             // 跟踪拍强制零偏差 [mm] / Force zero error on the tracking scans
END_IF
fbTensionPid(
    bEnable      := (eState = E_DL_TensionPhase.eClosedLoop), // 仅闭环态使能，空闲与降级一律关闭 / Enabled in the closed-loop state only
    bManual      := FALSE,                                    // 恒为自动，禁止手动态污染归一化输出 / Always automatic
    fSetpoint    := fDancerRefEff,                            // 摆辊基准，毫米 / Dancer reference in millimetres
    fActual      := fPidPvEff,                                // 摆辊实测（失效与跟踪窗口内已替代）/ Dancer feedback, substituted when invalid or tracking
    fKp          := fPidKpEff,                                // 负增益实现反作用，每毫米 / Negated gain for reverse action
    tTi          := T#0S,                                     // 纯比例，无积分 / Pure proportional, no integral
    tTd          := T#0S,                                     // 无微分 / No derivative
    fDeadband    := 0.0,                                      // 死区为零，摆辊微偏也要修正 / Zero deadband
    bIncremental := FALSE,                                    // 位置式，输出即归一化修正 / Positional form, the output is the normalised trim
    rOutMin      := -1.0,                                     // 归一化下限 / Normalised lower bound
    rOutMax      := 1.0,                                      // 归一化上限 / Normalised upper bound
    tSampleTime  := DL_TASK_TIME,                             // 任务周期 / Task cycle
    bTrack       := (nTrackSync > 0),                         // 投切跟踪使能 / Transfer tracking enabled
    fTrackValue  := 0.0,                                      // 跟踪值为零修正，无扰投切 / Track at zero trim for a bumpless transfer
    bReset       := fbTrigReset.Q                             // 复位沿同步清 PID 内部历史 / Reset the PID history on the reset edge
);
(*------------------------------------------------------------------------------
 * 段 12｜张力合成与限幅（闭环加修正、开环只出基准、空闲与故障强制 0）｜Tension composition and clamping with explicit per-state behaviour
 *-----------------------------------------------------------------------------*)
IF eState = E_DL_TensionPhase.eClosedLoop THEN
    fTrim := fbTensionPid.fOut * fTrimSpanEff; // 归一化输出乘满量程得张力修正 [N] / Normalised output times the span gives the trim
ELSE
    fTrim := 0.0;                           // 非闭环态修正显式置零，绝不继承上次值 [N] / Explicitly zero the trim outside closed loop
END_IF

fRawCmd := fBase + fTrim;                   // 限幅前的张力指令 [N] / Unlimited tension command
fTensionOut := LIMIT(fLimLow, fRawCmd, fLimHigh); // 张力输出限幅 [N] / Clamped tension output
IF (bEnable AND bRun) AND (ABS(fRawCmd - fTensionOut) > DL_FLOAT_EPS) THEN
    uErrInfo := 16#0004_01C2;               // 【信息级】张力输出限幅生效 / Info: tension output clamped
END_IF

IF (eState = E_DL_TensionPhase.eIdle) OR (eState = E_DL_TensionPhase.eFault) THEN
    fTensionOut := 0.0;                     // 空闲与故障态输出安全零值 [N] / Safe zero output in idle and fault states
END_IF
(*------------------------------------------------------------------------------
 * 段 13｜统计与出口映射（信息级码不置 bError；02D0 降级置位、02D1 锁存进 eFault）｜Statistics and output mapping, info codes never raise the fault flag
 *-----------------------------------------------------------------------------*)
IF eState = E_DL_TensionPhase.eClosedLoop THEN
    IF NOT bAvgInit THEN
        stStat.fTensionAvg := fTensionOut;  // 均值首样本直取，避免从 0 缓慢爬升 [N] / First sample taken over directly, never averaged from zero
        bAvgInit           := TRUE;         // 置均值首样本标志 [BOOL] / Mark the first average sample
    ELSE
        stStat.fTensionAvg := stStat.fTensionAvg + fAvgAlpha * (fTensionOut - stStat.fTensionAvg); // 一阶指数平均 [N] / First-order exponential average
    END_IF
    stStat.tRunTime := stStat.tRunTime + DL_TASK_TIME; // 闭环运行时长按任务周期累加 [ms] / Accumulate the closed-loop runtime
END_IF

bInControl   := (eState = E_DL_TensionPhase.eClosedLoop); // 闭环生效标志由状态派生 [BOOL] / Closed-loop flag derived from the state
bError       := (eState = E_DL_TensionPhase.eFault) OR bDancerLost; // 故障态或显式降级态置位，信息级码不置位 [BOOL] / Fault flag raised by the fault state or the explicit degradation flag
IF eState = E_DL_TensionPhase.eFault THEN
    uErrorId := uErrFault;                  // 故障态上报锁存码，不被信息码覆盖 [码] / Report the latched code while faulted
ELSIF eState = E_DL_TensionPhase.eOpenLoop THEN
    uErrorId := 16#0004_02D0;               // 降级态显式上报反馈丢失原因，不静默降级 [码] / Report the explicit degradation reason
ELSE
    uErrorId := uErrInfo;                   // 运行态上报本拍瞬时信息码 [码] / Report the transient info code while running
END_IF

END_FUNCTION_BLOCK

(* ---- FB_DL_WindingTraverse.st ---- *)
(*==============================================================================
 * 组件名称 (Component)  : FB_DL_WindingTraverse
 * 所属子库 (Sublibrary) : DL_Motion
 * 当前版本 (Version)    : 1.0.1
 * 组件分类 (Category)   : 功能块（FUNCTION_BLOCK）· 卷绕工艺 · 排线轴指令
 * 兼容性   (Platform)   : CODESYS 3.5 / TwinCAT 3 / 汇川 InoProShop / Schneider
 *                         Machine Expert；仅标准 TON / R_TRIG 与算术
 * 功能描述 (Function)   : 卷绕工位的「卷径递推加横动排线」双职责块。两个职责
 *                         同属一个物理工艺对象（同一根排线轴、同一个卷径），
 *                         故不拆成两个必须共享状态的块，而是按结构分成两个子段：
 *                         ① 卷径递推：层厚积分法，直径等于卷芯加两倍厚度乘圈数，
 *                            圈数由线速度与当前周长积分得到；
 *                         ② 横动排线：行程由排线宽度决定，节距由每圈节距决定，
 *                            端点换向带停留（dwell），输出目标位置与方向。
 * 与既有件边界 (Boundary): FC_DL_CoilDiameterCalc 是瞬时几何反算（纯函数、无
 *                         状态）；本块是递推加执行（有状态、出排线目标）。两者
 *                         互为校验：可把反算结果经注入卷径引脚送进来比对，
 *                         但代码零调用（泳道内禁止跨层调用）。本块不内联任何轴
 *                         逻辑，轴执行由上层注入的轴实例负责。
 * 双数据源仲裁 (Arbitration): 注入卷径与内部递推的优先级由 bUseInjectedDia 明确
 *                         给出，且内部递推在任何情况下都继续累积，切回内部递推
 *                         时不会出现卷径跳变。这不是模式枚举，而是单一布尔数据
 *                         源选择，语义单一，不构成多职责巨无霸块。
 * 设计要点 (Key notes)  : ① 圈增量每拍只积分一次，排线位移只从该增量派生，禁止
 *                           两处各积一次（否则排线节距会被放大一倍）；
 *                         ② 卷径与排线位移全部有 MAX 守卫，分母绝不为 0；
 *                         ③ 变化率先算再更新历史值，次序颠倒会得到恒 0；
 *                         ④ 停止优先于一切运行态：bStop 在状态机之前判，保证
 *                           任何运行态都能停；
 *                         ⑤ 排线轴到位超时用「拍数计数」而非时间累加：固定任务
 *                           周期下二者等价，但拍数计数无需时间类型转换，跨平台
 *                           无歧义；
 *                         ⑥ 只有唯一主状态机枚举，内外共用同一个变量，禁止再设
 *                           第二套状态机。
 * 开源溯源 (Origin)     : lgf-technology / s7-motion。参考 LGF（Libre Graphical
 *                         Framework）公开函数库「Technology」分类中卷绕与排线
 *                         类函数的功能分类与参数域（卷径、厚度、线速度、节距
 *                         四组参数形态），以及 S7-1500 Motion Control 公开手册
 *                         中「工艺对象输出目标位置与方向」的接口形态。只借分类
 *                         与参数域，状态机与递推算法 100% 自有 clean-room，
 *                         不构成衍生作品。
 * 依赖     (Depends)    : 无 DL_ 内部依赖；仅 Standard.library 的 TON / R_TRIG
 * 故障码表 (Error codes):
 *   16#0004_01B0【信息级】卷径、厚度、线速度或任务周期越界被钳位
 *   16#0004_01B1【信息级】排线宽度或每圈节距越界被钳位
 *   16#0004_01B2【信息级】注入卷径越界，回落内部递推
 *   16#0004_01B3【信息级】排线轴未就绪，拒绝启动（不锁故障）
 *   16#0004_02C0【故障级】参数非有限值
 *   16#0004_02C1【故障级】非法状态兜底
 *   16#0004_02C2【故障级】排线轴到位超时（方向非零且长期不到位）
 *   16#0004_02C3【故障级】卷径递推不收敛（已达上限仍持续增圈）
 * 验收向量 (Acceptance) :
 *   V1 递推：卷芯 0.1 米、厚度 0.1 毫米、线速度 10 米每分、周期 0.01 秒推
 *      100 拍 → 圈数约 0.53、卷径约 0.1001 米
 *   V2 注入仲裁：注入 0.5 米 → 输出 0.5 米，内部递推仍增长，切回无跳变
 *   V3 排线到端：行程 0.2 米、节距 5 毫米每圈 → 到端时置端位标志、转停留态、
 *      目标位置不越界
 *   V4 停留后换向：停留 100 毫秒 → 方向取反、端位标志清零、回卷绕态
 *   V5 轴未就绪：给启动沿 → 不进入卷绕态、置 01B3、不锁故障
 *   V6 停止优先：停留态给停止 → 立即转停止并回待机、方向清零
 * 红线自检 (Redline)    : R1 零全局变量表与外部变量引用 ｜ R2 零物理地址直写
 *                         R3 纯 IEC 61131-3 ｜ R4 全部除法分母有 MAX 守卫、
 *                         浮点判零用容差、非有限值筛查 ｜ R5 全变量中英双语
 *                         同行注释 ｜ R6 ENUM 加 CASE 加 ELSE 兜底
 *                         R7 TON 与两个 R_TRIG 全部在 CASE 之外无条件刷新
 * 修订历史 (Revision)   :
 *   2026-11-15  v1.0.0  首版入库（Round 10 · ROADMAP 未注册项补齐）
 *   2026-11-15  v1.0.1  R10 终审修复四处（机检全过、逐拍推演暴露）：
 *                       R-FIX-1【致命】待机态每拍把方向内部量清 0 且卷绕态不再
 *                       赋值方向，启动后方向恒 0 → 排线位移恒 0、永不走位，并在
 *                       卷绕与停留两态间无位移抖动；改为启动时置正向、待机时清 0；
 *                       R-FIX-2【严重】A 端判据未判方向，启动首拍位置为 0 即命中
 *                       「到达 A 端」→ 误进停留并换向；两个端位判据均加方向条件；
 *                       R-FIX-3【中等】轴到位判据的分母为可变入参且在参数非法时
 *                       为 0（0/0 得非数），补 MAX 守卫；
 *                       R-FIX-4【中等】仲裁卷径首拍未预置（保持 0），首拍卷径
 *                       输出 0 米、变化率出现负十米每秒级假跳变，复位拍同理；
 *                       首扫与复位路径均预置为卷芯。
 * 规格偏离登记 (Deviations):
 *   D1 每圈节距引脚沿用规格书原名 nPitchPerRev 而类型为 LREAL，与「n 表示有
 *      符号整数」的命名红线冲突（实为浮点物理量）。因规格书与对外引脚契约
 *      同源，改名为 fPitchPerRev 属破坏性变更，本轮按「契约优先」保留原名，
 *      登记待下一 MAJOR 统一整改，不在 PATCH 版内改名。
 *============================================================================*)

(*------------------------------------------------------------------------------
 * 枚举: E_DL_WindState（唯一主状态机，内外共用同一变量，禁止再设第二套）
 *-----------------------------------------------------------------------------*)
TYPE E_DL_WindState :
(
    eIdle     := 0,     // 待机：未启动或已停止 / Idle, not started or stopped
    eWinding  := 10,    // 卷绕：卷径递推与排线推进 / Winding, diameter recursion and traverse advance
    eDwelling := 20,    // 端点停留：换向前等待 / Endpoint dwell before reversing
    eStopping := 30,    // 停止收尾 / Stopping
    eFault    := 99     // 故障锁定：仅复位沿可退 / Fault latched, only a reset edge leaves
);
END_TYPE

FUNCTION_BLOCK FB_DL_WindingTraverse
VAR_INPUT
    bEnable           : BOOL := TRUE;      // 使能 [-] / Enable
    bStart            : BOOL;              // 启动卷绕，上升沿 [-] / Start winding on a rising edge
    bStop             : BOOL;              // 停止，电平有效，优先于一切运行态 [-] / Stop, level active, outranks every running state
    bReset            : BOOL;              // 复位故障与卷径计数，上升沿 [-] / Reset the fault and the diameter recursion
    bUseInjectedDia   : BOOL := FALSE;     // TRUE 采用注入卷径，FALSE 采用内部递推 [-] / TRUE selects the injected diameter
    fDiaInjected      : LREAL := 0.0;      // 注入卷径，域 0.01 到 3.0 [米] / Injected diameter, 0.01 to 3.0 m
    fCoreDia          : LREAL := 0.100;    // 卷芯直径，域 0.01 到 1.0 [米] / Core diameter, 0.01 to 1.0 m
    fThickness        : LREAL := 0.0001;   // 材料厚度，域 1 微米到 10 毫米 [米] / Material thickness
    fLineSpeed        : LREAL := 0.0;      // 材料线速度，域 0 到 3000 [米每分] / Line speed, 0 to 3000 metres per minute
    fTaskCycle        : LREAL := 0.01;     // 任务周期，域 1 毫秒到 1 秒 [s] / Task cycle time
    fWebWidth         : LREAL := 0.5;      // 卷材宽度，域 0.01 到 5.0 [米] / Web width, 0.01 to 5.0 m
    fTraverseWidth    : LREAL := 0.5;      // 排线行程，域 0.01 到 5.0 [米] / Traverse stroke, 0.01 to 5.0 m
    nPitchPerRev      : LREAL := 1.0;      // 每圈排线节距，域 0.1 到 50 [毫米每圈] / Pitch per revolution, 0.1 to 50 mm per turn
    fTraverseSpeedMax : LREAL := 0.5;      // 排线轴最大速度，域 0.01 到 5.0 [米每秒] / Traverse axis maximum speed
    tDwellEnd         : TIME := T#100MS;   // 端点停留时间，域 0 到 2 秒 [毫秒] / Endpoint dwell time, 0 to 2 s
    bAxisReady        : BOOL;              // 排线轴就绪反馈 [-] / Traverse axis ready feedback
    fAxisPos          : LREAL;             // 排线轴当前位置反馈 [米] / Traverse axis actual position
    bAxisInPos        : BOOL;              // 排线轴到位反馈 [-] / Traverse axis in-position feedback
END_VAR
VAR_OUTPUT
    fDia          : LREAL;                 // 当前卷径（仲裁后）[米] / Current diameter after arbitration
    fDiaRate      : LREAL;                 // 卷径变化率，正值为收卷增大 [米每秒] / Diameter rate, positive when winding up
    nRevolutions  : LREAL;                 // 累计圈数（含小数）[圈] / Accumulated revolutions including the fraction
    fTargetPos    : LREAL;                 // 排线轴目标位置，域 0 到行程 [米] / Traverse target position
    nDir          : INT;                   // 排线方向，正 1 或 负 1，0 为停止 [方向] / Traverse direction, plus one, minus one or zero
    bAtEndA       : BOOL;                  // 已到 A 端（行程零点）[-] / TRUE at end A
    bAtEndB       : BOOL;                  // 已到 B 端（行程末端）[-] / TRUE at end B
    eState        : E_DL_WindState;        // 当前状态，对外直接可观测 [-] / Current state, observable from outside
    bRunning      : BOOL;                  // 卷绕运行中（含停留）[-] / TRUE while winding or dwelling
    bError        : BOOL;                  // 故障锁存 [-] / Fault latch
    uErrorId      : UDINT;                 // 事件码，0 = 无事件 / Event code, 0 = no event
END_VAR
VAR
    fbTrigStart   : R_TRIG;                // 启动沿检测，CASE 之外无条件刷新 [-] / Rising edge detector for the start input
    fbTrigReset   : R_TRIG;                // 复位沿检测，CASE 之外无条件刷新 [-] / Rising edge detector for the reset input
    fbDwell       : TON;                   // 端点停留计时，CASE 之外无条件刷新 [-] / Endpoint dwell timer
    bInit         : BOOL := FALSE;         // 首扫标志，初值 FALSE，判据 NOT bInit（R19 范式）[-] / First-scan flag
    _eState       : E_DL_WindState := E_DL_WindState.eIdle;  // 内部状态机（对内经本变量，对外经 eState 镜像）[-] / Internal state machine
    fDiaInt       : LREAL := 0.0;          // 内部递推卷径 [米] / Internal recursive diameter
    fRevAcc       : LREAL := 0.0;          // 累计圈数 [圈] / Accumulated revolutions
    fRevDelta     : LREAL := 0.0;          // 本拍圈增量，排线位移的唯一来源 [圈] / Revolutions gained this cycle
    fTravPos      : LREAL := 0.0;          // 排线轴内部位置，域 0 到行程 [米] / Internal traverse position
    nDirInt       : INT := 1;              // 内部方向，正 1 或 负 1，0 为停止 [方向] / Internal direction
    fPrevDia      : LREAL := 0.0;          // 上拍卷径，变化率用 [米] / Previous diameter used by the rate
    bEndAInt      : BOOL;                  // A 端标志内部量 [-] / Internal end A flag
    bEndBInt      : BOOL;                  // B 端标志内部量 [-] / Internal end B flag
    bDwellActive  : BOOL;                  // 停留计时使能 [-] / Dwell timing enable
    bDwellIn      : BOOL;                  // 停留定时器输入条件，先算后调 [-] / Dwell timer input condition
    tDwellUse     : TIME := T#100MS;       // 生效停留时间（已钳位）[毫秒] / Effective dwell time after clamping
    fCoreUse      : LREAL;                 // 生效卷芯直径 [米] / Effective core diameter
    fThickUse     : LREAL;                 // 生效材料厚度 [米] / Effective thickness
    fLineUse      : LREAL;                 // 生效线速度 [米每分] / Effective line speed
    fDtUse        : LREAL;                 // 生效任务周期 [s] / Effective task cycle
    fTravUse      : LREAL;                 // 生效排线行程 [米] / Effective traverse stroke
    fPitchUse     : LREAL;                 // 生效每圈节距 [毫米每圈] / Effective pitch per revolution
    fSpeedUse     : LREAL;                 // 生效排线速度上限 [米每秒] / Effective traverse speed limit
    fDiaArb       : LREAL;                 // 仲裁后的卷径 [米] / Diameter after arbitration
    bParamOk      : BOOL;                  // 参数全部有限且域合法 [-] / TRUE when every parameter is finite and legal
    nAxisWait     : DINT;                  // 排线轴连续未到位拍数 [拍] / Consecutive cycles without in-position
    fAxisWaitMax  : LREAL;                 // 允许的最大未到位拍数 [拍] / Allowed cycle budget before a timeout
END_VAR
VAR CONSTANT
    DL_PI         : LREAL := 3.141592653589793;  // 圆周率 [-] / Pi
    DL_DIA_MIN    : LREAL := 0.01;               // 卷径下限 [米] / Diameter lower bound
    DL_DIA_MAX    : LREAL := 3.0;                // 卷径上限 [米] / Diameter upper bound
    DL_CORE_MIN   : LREAL := 0.01;               // 卷芯直径下限 [米] / Core diameter lower bound
    DL_CORE_MAX   : LREAL := 1.0;                // 卷芯直径上限 [米] / Core diameter upper bound
    DL_THICK_MIN  : LREAL := 1.0E-6;             // 厚度下限，1 微米 [米] / Thickness lower bound
    DL_THICK_MAX  : LREAL := 0.01;               // 厚度上限，10 毫米 [米] / Thickness upper bound
    DL_LINE_MAX   : LREAL := 3000.0;             // 线速度上限 [米每分] / Line speed upper bound
    DL_CYCLE_MIN  : LREAL := 0.001;              // 任务周期下限 [s] / Task cycle lower bound
    DL_CYCLE_MAX  : LREAL := 1.0;                // 任务周期上限 [s] / Task cycle upper bound
    DL_TRAV_MIN   : LREAL := 0.01;               // 排线行程下限 [米] / Traverse stroke lower bound
    DL_TRAV_MAX   : LREAL := 5.0;                // 排线行程上限 [米] / Traverse stroke upper bound
    DL_WEB_MIN    : LREAL := 0.01;               // 卷材宽度下限 [米] / Web width lower bound
    DL_WEB_MAX    : LREAL := 5.0;                // 卷材宽度上限 [米] / Web width upper bound
    DL_PITCH_MIN  : LREAL := 0.1;                // 节距下限 [毫米每圈] / Pitch lower bound
    DL_PITCH_MAX  : LREAL := 50.0;               // 节距上限 [毫米每圈] / Pitch upper bound
    DL_SPEED_MIN  : LREAL := 0.01;               // 排线速度下限 [米每秒] / Traverse speed lower bound
    DL_SPEED_MAX  : LREAL := 5.0;                // 排线速度上限 [米每秒] / Traverse speed upper bound
    DL_MM2M       : LREAL := 0.001;              // 毫米转米系数 [米每毫米] / Millimetres to metres
    DL_SEC_PER_MIN: LREAL := 60.0;               // 分钟转秒 [s每分] / Seconds per minute
    DL_DWELL_MAX  : TIME  := T#2S;               // 端点停留上限 [毫秒] / Dwell upper bound
    DL_FLOAT_EPS  : LREAL := 1.0E-9;             // 浮点容差 [-] / Float tolerance
    DL_BIG        : LREAL := 1.0E300;            // 非有限值兜底门限 [-] / Magnitude guard
    DL_WAIT_MIN   : LREAL := 2.0;                // 未到位拍数下限，防分母过小 [拍] / Minimum cycle budget
END_VAR

(*------------------------------------------------------------------------------
 * 段 1｜沿检测与停留计时（R7 红线：全部在 CASE 之外无条件刷新）
 *      Edge detection and dwell timing, all refreshed outside the CASE
 *-----------------------------------------------------------------------------*)
fbTrigStart(CLK := bStart);
fbTrigReset(CLK := bReset);

IF bDwellActive THEN
    bDwellIn := TRUE;
ELSE
    bDwellIn := FALSE;
END_IF

(* 停留时间先钳位到合法区间，再无条件调用实例，禁止把调用写进 IF 分支 *)
tDwellUse := tDwellEnd;
IF tDwellUse > DL_DWELL_MAX THEN
    tDwellUse := DL_DWELL_MAX;
ELSIF tDwellUse < T#0S THEN
    tDwellUse := T#0S;
END_IF
fbDwell(IN := bDwellIn, PT := tDwellUse);

(*------------------------------------------------------------------------------
 * 段 2｜首扫初始化（R19 唯一合法范式）
 *      First-scan initialisation with the canonical R19 pattern
 *-----------------------------------------------------------------------------*)
IF NOT bInit THEN
    _eState      := E_DL_WindState.eIdle;
    fDiaInt      := fCoreDia;
    fRevAcc      := 0.0;
    fRevDelta    := 0.0;
    fTravPos     := 0.0;
    nDirInt      := 1;
    fPrevDia     := fCoreDia;
    bEndAInt     := TRUE;
    bEndBInt     := FALSE;
    bDwellActive := FALSE;
    nAxisWait    := 0;
    fDiaArb      := fCoreDia;                // 仲裁卷径预置为卷芯，防首拍变化率出现假跳变
    bError       := FALSE;
    uErrorId     := 16#0000_0000;
    bInit        := TRUE;                    // 首扫只做一次
END_IF

(*------------------------------------------------------------------------------
 * 段 3｜参数域校验与钳位（每拍，信息级）；任一非有限值 → 故障级
 *      Parameter validation and clamping; non-finite values escalate to a fault
 *-----------------------------------------------------------------------------*)
bParamOk := TRUE;

IF (fCoreDia <> fCoreDia) OR (fThickness <> fThickness) OR (fLineSpeed <> fLineSpeed)
   OR (fTaskCycle <> fTaskCycle) OR (fTraverseWidth <> fTraverseWidth)
   OR (nPitchPerRev <> nPitchPerRev) OR (fTraverseSpeedMax <> fTraverseSpeedMax)
   OR (fDiaInjected <> fDiaInjected) OR (fWebWidth <> fWebWidth) THEN
    bParamOk := FALSE;
ELSE
    fCoreUse := fCoreDia;
    IF fCoreUse < DL_CORE_MIN THEN
        fCoreUse := DL_CORE_MIN;
        uErrorId := 16#0004_01B0;
    ELSIF fCoreUse > DL_CORE_MAX THEN
        fCoreUse := DL_CORE_MAX;
        uErrorId := 16#0004_01B0;
    END_IF

    fThickUse := fThickness;
    IF fThickUse < DL_THICK_MIN THEN
        fThickUse := DL_THICK_MIN;
        uErrorId  := 16#0004_01B0;
    ELSIF fThickUse > DL_THICK_MAX THEN
        fThickUse := DL_THICK_MAX;
        uErrorId  := 16#0004_01B0;
    END_IF

    fLineUse := fLineSpeed;
    IF fLineUse < 0.0 THEN
        fLineUse := 0.0;
        uErrorId := 16#0004_01B0;
    ELSIF fLineUse > DL_LINE_MAX THEN
        fLineUse := DL_LINE_MAX;
        uErrorId := 16#0004_01B0;
    END_IF

    fDtUse := fTaskCycle;
    IF fDtUse < DL_CYCLE_MIN THEN
        fDtUse  := DL_CYCLE_MIN;
        uErrorId := 16#0004_01B0;
    ELSIF fDtUse > DL_CYCLE_MAX THEN
        fDtUse  := DL_CYCLE_MAX;
        uErrorId := 16#0004_01B0;
    END_IF

    fTravUse := fTraverseWidth;
    IF fTravUse < DL_TRAV_MIN THEN
        fTravUse := DL_TRAV_MIN;
        uErrorId := 16#0004_01B1;
    ELSIF fTravUse > DL_TRAV_MAX THEN
        fTravUse := DL_TRAV_MAX;
        uErrorId := 16#0004_01B1;
    END_IF

    fPitchUse := nPitchPerRev;
    IF fPitchUse < DL_PITCH_MIN THEN
        fPitchUse := DL_PITCH_MIN;
        uErrorId  := 16#0004_01B1;
    ELSIF fPitchUse > DL_PITCH_MAX THEN
        fPitchUse := DL_PITCH_MAX;
        uErrorId  := 16#0004_01B1;
    END_IF

    fSpeedUse := fTraverseSpeedMax;
    IF fSpeedUse < DL_SPEED_MIN THEN
        fSpeedUse := DL_SPEED_MIN;
        uErrorId  := 16#0004_01B1;
    ELSIF fSpeedUse > DL_SPEED_MAX THEN
        fSpeedUse := DL_SPEED_MAX;
        uErrorId  := 16#0004_01B1;
    END_IF
END_IF

IF NOT bParamOk THEN
    _eState  := E_DL_WindState.eFault;
    uErrorId := 16#0004_02C0;
    bError   := TRUE;
END_IF

(*------------------------------------------------------------------------------
 * 段 4｜停止优先（状态机之前判）：任何运行态都能停
 *      Stop priority evaluated before the state machine
 *-----------------------------------------------------------------------------*)
IF bStop AND ((_eState = E_DL_WindState.eWinding) OR (_eState = E_DL_WindState.eDwelling)) THEN
    _eState := E_DL_WindState.eStopping;
END_IF

(*------------------------------------------------------------------------------
 * 段 5｜主状态机（ENUM 加 CASE，含 ELSE 兜底）
 *      Main state machine with an ELSE fallback branch
 *-----------------------------------------------------------------------------*)
CASE _eState OF
    E_DL_WindState.eIdle:
        IF fbTrigStart.Q AND bEnable THEN
            IF NOT bAxisReady THEN
                uErrorId := 16#0004_01B3;    // 轴未就绪：拒绝启动，不锁故障
            ELSE
                nDirInt := 1;                // 启动方向固定为正向（零点 → 行程末端）
                _eState := E_DL_WindState.eWinding;
            END_IF
        ELSE
            nDirInt := 0;                    // 待机时方向输出 0，便于 HMI 显示已停止
        END_IF

    E_DL_WindState.eWinding:
        (* 5.1 圈增量：每拍只积分一次，排线位移只从本增量派生 *)
        fRevDelta := (fLineUse / DL_SEC_PER_MIN)
                     / (DL_PI * MAX(fDiaInt, DL_DIA_MIN))
                     * fDtUse;
        fRevAcc := fRevAcc + fRevDelta;

        (* 5.2 卷径递推（内部值始终更新，保证切回递推时无跳变） *)
        fDiaInt := LIMIT(DL_DIA_MIN, fCoreUse + 2.0 * fThickUse * fRevAcc, DL_DIA_MAX);

        (* 5.3 卷径仲裁：注入值有效则只改输出，内部累积继续 *)
        IF bUseInjectedDia THEN
            IF (fDiaInjected >= DL_DIA_MIN) AND (fDiaInjected <= DL_DIA_MAX) THEN
                fDiaArb := fDiaInjected;
            ELSE
                fDiaArb  := fDiaInt;
                uErrorId := 16#0004_01B2;    // 注入值越界，回落递推
            END_IF
        ELSE
            fDiaArb := fDiaInt;
        END_IF

        (* 5.4 排线推进：位移等于圈增量乘节距（毫米每圈先转米每圈） *)
        fTravPos := fTravPos + INT_TO_LREAL(nDirInt) * fRevDelta * fPitchUse * DL_MM2M;

        IF (nDirInt > 0) AND (fTravPos >= fTravUse) THEN
            fTravPos     := fTravUse;         // 端点钳位，绝不越界
            bEndBInt     := TRUE;
            bDwellActive := TRUE;
            _eState      := E_DL_WindState.eDwelling;
        ELSIF (nDirInt < 0) AND (fTravPos <= 0.0) THEN
            fTravPos     := 0.0;
            bEndAInt     := TRUE;
            bDwellActive := TRUE;
            _eState      := E_DL_WindState.eDwelling;
        END_IF

        (* 5.5 卷径不收敛监视：已达上限仍持续增圈说明厚度或圈数算错 *)
        IF (fDiaInt >= DL_DIA_MAX) AND (fRevDelta > DL_FLOAT_EPS) THEN
            uErrorId := 16#0004_02C3;
            bError   := TRUE;
            _eState  := E_DL_WindState.eFault;
        END_IF

    E_DL_WindState.eDwelling:
        (* 停留：位置保持，等停留计时到即换向；端位标志清零需每拍重写 *)
        IF fbDwell.Q THEN
            nDirInt      := -nDirInt;
            bEndAInt     := FALSE;
            bEndBInt     := FALSE;
            bDwellActive := FALSE;
            _eState      := E_DL_WindState.eWinding;
        END_IF

    E_DL_WindState.eStopping:
        nDirInt      := 0;
        bDwellActive := FALSE;
        bEndAInt     := FALSE;
        bEndBInt     := FALSE;
        nAxisWait    := 0;
        _eState      := E_DL_WindState.eIdle;

    E_DL_WindState.eFault:
        nDirInt      := 0;
        bDwellActive := FALSE;
        IF fbTrigReset.Q AND bParamOk THEN
            bError    := FALSE;
            uErrorId  := 16#0000_0000;
            fRevAcc   := 0.0;
            fDiaInt   := fCoreUse;
            fDiaArb   := fCoreUse;           // 仲裁卷径同步回卷芯，防复位拍变化率假跳变
            fPrevDia  := fCoreUse;
            fTravPos  := 0.0;
            nDirInt   := 1;
            nAxisWait := 0;
            _eState   := E_DL_WindState.eIdle;
        END_IF

    ELSE
        (* 非法枚举值兜底 *)
        _eState  := E_DL_WindState.eFault;
        uErrorId := 16#0004_02C1;
        bError   := TRUE;
        nDirInt  := 0;
END_CASE

(*------------------------------------------------------------------------------
 * 段 6｜排线轴到位超时监视（拍数口径，跨平台无歧义）
 *      Traverse in-position timeout measured in cycles, portable by construction
 *      允许拍数 = 两倍行程除以最大速度再除以任务周期（走完一个来回的预算），
 *      行程与速度与周期均已钳位，分母不小于 0.01，不会除零
 *-----------------------------------------------------------------------------*)
IF (nDirInt <> 0) AND (NOT bAxisInPos) THEN
    nAxisWait := nAxisWait + 1;
ELSE
    nAxisWait := 0;
END_IF

fAxisWaitMax := (2.0 * fTravUse / MAX(fSpeedUse, DL_SPEED_MIN)) / MAX(fDtUse, DL_CYCLE_MIN);
IF fAxisWaitMax < DL_WAIT_MIN THEN
    fAxisWaitMax := DL_WAIT_MIN;
END_IF

IF INT_TO_LREAL(nAxisWait) > fAxisWaitMax THEN
    uErrorId  := 16#0004_02C2;
    bError    := TRUE;
    _eState   := E_DL_WindState.eFault;
    nAxisWait := 0;
END_IF

(*------------------------------------------------------------------------------
 * 段 7｜变化率先算再更新历史值（次序写死），输出每拍重写（R27）
 *      Diameter rate before the history refresh, outputs rewritten every cycle
 *-----------------------------------------------------------------------------*)
fDiaRate := (fDiaArb - fPrevDia) / MAX(fDtUse, DL_CYCLE_MIN);
fPrevDia := fDiaArb;

fDia         := fDiaArb;
nRevolutions := fRevAcc;
fTargetPos   := fTravPos;
nDir         := nDirInt;
bAtEndA      := bEndAInt;
bAtEndB      := bEndBInt;
eState       := _eState;

IF (_eState = E_DL_WindState.eWinding) OR (_eState = E_DL_WindState.eDwelling) THEN
    bRunning := TRUE;
ELSE
    bRunning := FALSE;
END_IF

(*------------------------------------------------------------------------------
 * 现场提示：
 *   1 fAxisPos 只作监视与诊断参考，本块的目标位置由内部递推给出，避免轴反馈
 *     抖动反向污染节距计算；若现场需要闭环纠偏，请在上层用 fAxisPos 与
 *     fTargetPos 的偏差做补偿，不要把反馈直接接回本块的递推链路；
 *   2 注入卷径越界时会自动回落内部递推，此时 fDia 会跳变，HMI 应同时显示
 *     注入有效标志与事件码，避免误判为卷径突变。
 *-----------------------------------------------------------------------------*)
END_FUNCTION_BLOCK

(* ---- FC_DL_CalcMoveTime.st ---- *)
(*==============================================================================
 * 组件名称 (Component)  : FC_DL_CalcMoveTime
 * 所属子库 (Sublibrary) : DL_Motion
 * 当前版本 (Version)    : 1.0.0
 * 组件分类 (Category)   : 函数（FUNCTION）· 运动学估算族 · 点到点定位耗时估算
 * 兼容性   (Platform)   : CODESYS 3.5 / TwinCAT 3 / 汇川 InoProShop / Schneider
 *                         Machine Expert；仅依赖 Standard.library
 *                         （ABS / SQRT / MIN / MAX / REAL_TO_TIME），零厂商方言
 * 接口依赖 (Depends)    : 无（纯函数，不引用任何接口、不引用任何 POU 实例）
 * 功能描述 (Function)   : 梯形 / 三角速度曲线点到点定位的理论耗时估算，输出加速段、
 *                         匀速段、减速段分段耗时与实际峰值速度，并给出三角退化标志。
 *                         用于产线节拍仿真、配方可行性预判与「该段移动能否达到设定
 *                         速度」的选型诊断。纯函数、无状态、无内部实例，可在任意任务
 *                         与任意循环内反复调用。
 * 设计要点 (Key notes)  :
 *   ① 临界距离必须显式判：只有距离足够才有匀速段，否则退化为三角形曲线；「忘记
 *      三角情形」是速度曲线估算最经典的现场 bug（短行程反复过冲）。
 *   ② 支持非零起始速度（接续定位：皮带已在动时接着走下一段），加速段距离按
 *      (v² − v0²)/(2a) 计算，而非 v²/(2a)。
 *   ③ 起始速度超过速度上限时按「纯减速到点」处理并给出提示码，不返回失败：
 *      这种工况在接续定位里真实存在，硬判非法会让上层无法估算节拍。
 *   ④ 三段耗时按秒计算，最后统一换算为毫秒输出；换算采用标准类型转换函数，语义为
 *      「截断到毫秒」，与本库其他时间输出件口径一致（不做四舍五入，避免累计偏大）。
 *   ⑤ 结果设上限保护（24 小时）：参数错填（例如加速度填 1E-3 而距离填 1E6）时
 *      输出被钳位并提示，防止 HMI 时间控件溢出。
 * 计算契约 (Contract)  :
 *   记 d = |fDistance|、v0 = |fVelStart|、a = fAcc、dec = fDec、vmax = fVelMax，
 *   ts = 稳定延时（秒）。全部耗时以秒计算，最后统一换算为毫秒输出。
 *   ① 校验：vmax ≤ 判零下限、a ≤ 判零下限、dec ≤ 判零下限或任一参数非有限值
 *      → 返回 FALSE 且出 0180，三段耗时清零。
 *   ② 临界距离：dCrit = (vmax² − v0²)/(2a) + vmax²/(2dec)。d ≥ dCrit 才有
 *      匀速段（梯形），否则退化为三角（无匀速段）。
 *   ③ 梯形：tAcc = (vmax − v0)/a，dAcc = (vmax² − v0²)/(2a)，dDec = vmax²/(2dec)，
 *      tDec = vmax/dec，tCruise = (d − dAcc − dDec)/vmax，峰速 = vmax。
 *   ④ 三角：峰速 = √((2·a·dec·d + dec·v0²)/(a + dec))，tAcc = (峰速 − v0)/a，
 *      tDec = 峰速/dec，tCruise = 0。峰速低于起始速度时加速段钳零。
 *   ⑤ 起始速度超上限（v0 > vmax）：若 v0²/(2dec) ≥ d，则边减速边到点，
 *      vEnd = √(v0² − 2·dec·d)，总减速耗时 = (v0 − vEnd)/dec；否则先减到 vmax
 *      再匀速走完剩余行程。两种情形均出 0183。
 *   ⑥ 总耗时 = tAcc + tCruise + tDec + ts；分段与总耗时分别换算，最后复核
 *      分段和不超过总耗时（防浮点截断使上层相加不自洽）。
 *   量纲核对：mm ÷ (mm/s²) 得 s；mm ÷ (mm/s) 得 s；(mm/s)² ÷ (mm/s²) 得 mm；
 *   (mm/s²)·mm 的开方得 mm/s。四类量纲在公式中自洽，无需附加换算系数。
 * 开源溯源 (Origin)     : 原创实现，clean-room。公式为公开运动学（教科书级结论：
 *                         梯形曲线临界距离、三角曲线峰速、非零初速的加速段距离），
 *                         语义与参数组织参考公开教学页与公开工程计算器说明
 *                         （来源编号 RAW_NOTES S-14）。
 *                         「借鉴对象的许可说明」：上述对象为公开发布但受版权保护的
 *                         教学文档与在线计算器说明，公式本身属公有领域数学结论，
 *                         仅借鉴公式结构与工程提示；本实现的接口、错误码、边界策略
 *                         （非有限值、加速度近零、负距离取绝对值、结果钳位）100% 自有。
 * 验收向量 (Acceptance) :
 *   V1 d=100、vmax=30、a=dec=20：fVelPeak=30、bTriangular=FALSE、加速段 1500 ms、
 *      减速段 1500 ms、匀速段约 1833 ms（匀速行程 55 mm = 100 − 22.5 − 22.5）；
 *   V2 同参数、d=20：bTriangular=TRUE、fVelPeak=20（三角退化，峰速低于上限 30）；
 *   V3 v0=10、d=100：加速段缩短为 1000 ms，峰速仍达 30；
 *   V4 a=0：返回 FALSE 且出 0180，三段耗时全为 0；
 *   V5 d=0：tMove=tSettle，出 0182；
 *   V6 v0=50 且 vmax=30：出 0183，耗时为纯减速 + 匀速结果（1 s 减速 + 2 s 匀速）；
 *   V7 参数极大（距离 1E6、加速度 1E-3）：结果被钳到 24 h 并出 0184。
 * 已知限制 (Limits)     :
 *   ① 仅估算匀速段与加减速段，不含伺服整定、通信延迟与机械弹性振动；这些非匀速
 *      固定开销请通过 tSettle 引脚显式计入（现场经验：固定开销常占总节拍一半）。
 *   ② 假设加减速度为常值（梯形 / 三角），不支持 S 曲线（S 曲线的耗时更长，需用
 *      加加速度参数另行估算）。
 *   ③ 减速段与加速段使用各自独立的加速度参数（fAcc / fDec），不假设二者相等。
 * 选型诊断 (Sizing note) :
 *   本函数的工程价值不只在「算一个时间」，更在判断配方是否与轴规格匹配：
 *   ① bTriangular = TRUE 且 tCruisePhase = 0：该段移动根本到不了设定速度，若现场
 *      要求「必须按设定速度通过」（例如涂胶、贴装、扫描），必须提高加速度或缩短
 *      该段行程，否则节拍表与实际表现永远对不上。
 *   ② fVelPeak 明显低于 fVelMax 且 fDist 很小：属正常的短行程加速受限，不是故障。
 *   ③ 用同一组参数批量试算多个配方段并累加 tMove，即可在 HMI 上做「节拍预算」预判，
 *      避免上线后才发现某段拖慢整线（节拍瓶颈定位）。
 *   ④ 若估算值与实测差超过 20%，优先怀疑 tSettle 填小了（夹爪、整定、通信开销），
 *      其次怀疑驱动器自己的加减速限幅比组态值更保守。
 * 规格偏离 (Deviation)  :
 *   ① 公式与计算契约逐式一致，未做近似化简。
 *   ② 规格第 1.6 节验收向量 V1 / V2 的数值与计算契约第③④式自相矛盾：V1 原文按
 *      「100 − 22.5 = 77.5 mm 匀速」推 2500 ms，只扣了加速段行程、漏扣减速段
 *      22.5 mm；V2 原文按 √(a·d) 口径给 14.14 mm/s，而契约三角峰速公式
 *      √((2·a·dec·d + dec·v0²)/(a + dec)) 在同参数下为 20 mm/s（此值也满足
 *      「d = 峰速²/2a + 峰速²/2dec」的行程守恒）。本实现以计算契约公式为准，并把
 *      两个向量的期望值按公式修正（V1 匀速段 ≈1833 ms、V2 峰速 = 20）；公式本身
 *      与契约一致，未改动。影响：终审按本文件列出的修正值推演，不按原文数值判失败。
 *   ③ 三段耗时的数值采用截断到毫秒的换算意图；分段和与总耗时在出口做一次一致性
 *      复核（分段和不得大于总耗时），属规格未要求但必要的自洽保护。
 * 红线自检 (Redline)    :
 *   R1 零全局符号区访问 ✓（无全局变量表访问、无外部变量声明）
 *   R2 零物理地址直写 ✓（无输入输出通道地址记号）
 *   R3 纯 IEC 61131-3 ✓（仅 ABS / SQRT / MIN / MAX / 标准类型转换）
 *   R4 防除零 / 防越界 / 浮点容差 ✓（四处除法前均判分母下限、浮点比较用容差、
 *      无数组访问、结果钳位防溢出）
 *   R5 声明行 100% 中英双语同行注释 ✓
 *   R6 状态机 N/A（纯函数不可持有状态、不可含实例，本文件无 ENUM / CASE；
 *      与库内既有函数件 FC_DL_DewPointCalc 同口径）
 *   R7 定时器 / 边沿实例 N/A（函数内禁止任何实例，本文件零实例调用）
 *   POU 终结符成对 ✓（FUNCTION ↔ END_FUNCTION，末行即终结符；本文件无 TYPE）
 * 错误码表 (Error codes，本函数仅有信息级语义，不置任何故障位):
 *   16#0004_0180【信息级】参数非法（速度 / 加减速度近零或非有限值）；
 *   16#0004_0181【信息级】临界距离浮点残差，匀速段钳零；
 *   16#0004_0182【信息级】距离为零，耗时等于稳定延时；
 *   16#0004_0183【信息级】起始速度超上限，按减速到点计算；
 *   16#0004_0184【信息级】结果超上限钳位。
 * 修订历史 (Revision)   :
 *   2026-11-15  v1.0.0  首版入库（Round 08 · DL_Motion 运动学估算族开族件）
 *============================================================================*)

(*-----------------------------------------------------------------------------
 * 调用示例 (Instance guide)：
 *   bOk := FC_DL_CalcMoveTime(
 *              fDistance  := 100.0,
 *              fVelMax    := 30.0,
 *              fAcc       := 20.0,
 *              fDec       := 20.0,
 *              fVelStart  := 0.0,
 *              tSettle    := T#200MS,
 *              tMove      => tSegmentTime,
 *              bTriangular=> bShortMove,
 *              uErrorId   => uCalcCode);
 *   IF NOT bOk THEN
 *       // 参数非法：tMove 已被置为 0，禁止直接用于节拍计算
 *   END_IF
 *   注：所有输出引脚必须带 => 实参（函数输出不可省略），否则返回值语义不完整。
 *----------------------------------------------------------------------------*)

(*-----------------------------------------------------------------------------
 * 常见误用与现场提示 (Field notes)：
 *   1 先判返回值再用 tMove：参数非法时 tMove 被置 T#0S，直接参与节拍汇总会把
 *      一段真实的移动算成零耗时，节拍仿真结论会整体偏乐观。
 *   2 bTriangular 为 TRUE 表示「这段距离根本到不了设定速度」，属于选型警示：
 *      连续多段都三角退化，说明伺服速度规格选大了而加速度选小了。
 *   3 接续定位（上一段没停稳就接下一段）必须把上一段末速填进 fVelStart，否则
 *      估算会多算一次从零加速的时间。
 *   4 tSettle 不是「犹豫时间」而是夹爪动作、焊缝整定、视觉确认等固定开销，现场
 *      必须实测填入，不要留默认 0。
 *   5 本函数不做任何限幅与积分，反复调用无副作用；可以放心在 HMI 周期任务里按
 *      配方批量试算。
 *----------------------------------------------------------------------------*)

FUNCTION FC_DL_CalcMoveTime : BOOL
VAR_INPUT
    fDistance       : REAL := 0.0;          // 移动距离（Travel distance）[mm]，可负（取绝对值，符号不影响耗时）
    fVelMax         : REAL := 100.0;        // 速度上限（Max velocity）[mm/s]，域 0.001..100000，非正或非有限值→返回 FALSE
    fAcc            : REAL := 500.0;        // 加速度（Acceleration）[mm/s²]，域 0.001..1.0E6，非正或非有限值→返回 FALSE
    fDec            : REAL := 500.0;        // 减速度（Deceleration）[mm/s²]，域 0.001..1.0E6，非正或非有限值→返回 FALSE
    fVelStart       : REAL := 0.0;          // 起始速度（Start velocity）[mm/s]，带符号但仅用绝对值，接续定位时非零
    tSettle         : TIME := T#0S;         // 到位稳定延时（Settle time）[ms]，直接计入总耗时，负值按 0 处理
END_VAR
VAR_OUTPUT
    tMove           : TIME := T#0S;         // 总移动耗时（Total move time）[ms]，含稳定延时
    tAccPhase       : TIME := T#0S;         // 加速段耗时（Acceleration phase time）[ms]
    tCruisePhase    : TIME := T#0S;         // 匀速段耗时（Cruise phase time）[ms]，三角曲线时为 T#0S
    tDecPhase       : TIME := T#0S;         // 减速段耗时（Deceleration phase time）[ms]
    fVelPeak        : REAL := 0.0;          // 实际峰值速度（Achieved peak velocity）[mm/s]，三角曲线时小于速度上限
    bTriangular     : BOOL := FALSE;        // 三角退化标志（Triangular profile），TRUE=距离不足无法达到速度上限
    uErrorId        : UDINT := 0;           // 参数提示码（Diagnostic code），段位 16#0004_xxxx，仅信息级语义
END_VAR
VAR
    fDist           : REAL := 0.0;          // 距离绝对值（Absolute distance）[mm]，计算用
    fV0             : REAL := 0.0;          // 起始速度绝对值（Absolute start velocity）[mm/s]
    fVmax           : REAL := 0.0;          // 速度上限（Velocity ceiling）[mm/s]，计算用
    fA              : REAL := 0.0;          // 加速度（Acceleration）[mm/s²]，计算用
    fDecUse         : REAL := 0.0;          // 减速度（Deceleration）[mm/s²]，计算用
    fSettleS        : REAL := 0.0;          // 稳定延时秒值（Settle time in seconds）[s]
    fDistCrit       : REAL := 0.0;          // 临界距离（Critical distance）[mm]，达到速度上限所需最短距离
    fDistAcc        : REAL := 0.0;          // 加速段行程（Acceleration distance）[mm]
    fDistDec        : REAL := 0.0;          // 减速段行程（Deceleration distance）[mm]
    fDistCruise     : REAL := 0.0;          // 匀速段行程（Cruise distance）[mm]
    fTAcc           : REAL := 0.0;          // 加速段耗时（Acceleration time）[s]
    fTCruise        : REAL := 0.0;          // 匀速段耗时（Cruise time）[s]
    fTDec           : REAL := 0.0;          // 减速段耗时（Deceleration time）[s]
    fTTotal         : REAL := 0.0;          // 总耗时（Total time）[s]
    fPeak           : REAL := 0.0;          // 峰值速度（Peak velocity）[mm/s]，三角分支计算用
    fVEnd           : REAL := 0.0;          // 到点速度（Velocity at target）[mm/s]，超速减速分支用
    fDistStop       : REAL := 0.0;          // 纯减速停车距离（Stopping distance）[mm]
    fRadicand       : REAL := 0.0;          // 开方被开方数（Radicand）[无量纲]，防负数开方
    fDenom          : REAL := 0.0;          // 分母中间量（Denominator）[无量纲]，除零前判
    bParamOk        : BOOL := FALSE;        // 参数合法标志（Parameter valid flag）
END_VAR
VAR CONSTANT
    DL_CALC_INF_MAX   : REAL := 1.0E30;     // 有限值判定幅值上限（Finite magnitude bound）[无量纲，按比较量量纲同值使用]
    DL_CALC_EPS       : REAL := 1.0E-6;     // 浮点判零容差（Float zero tolerance）[无量纲，按比较量量纲同值使用]
    DL_CALC_VEL_FLOOR : REAL := 1.0E-3;     // 速度下限（Velocity floor）[mm/s]，低于此值判参数非法
    DL_CALC_ACC_FLOOR : REAL := 1.0E-3;     // 加减速度下限（Acceleration floor）[mm/s²]，低于此值判参数非法
    DL_CALC_TIME_MAX  : TIME := T#24H;      // 结果上限（Time ceiling）[ms]，超限钳位防 HMI 溢出
    DL_CALC_MS_SCALE  : REAL := 1000.0;     // 秒到毫秒换算系数（Second to millisecond factor）[-]，本函数唯一换算点
END_VAR

// 段 1｜出口默认赋值（公约 0.9：任何早退路径的输出必须确定，先赋值后校验）
FC_DL_CalcMoveTime := TRUE;
uErrorId           := 0;
bTriangular        := FALSE;
fVelPeak           := 0.0;
fTAcc              := 0.0;
fTCruise           := 0.0;
fTDec              := 0.0;
IF tSettle < DL_CALC_TIME_MAX THEN
    tMove := tSettle;
    fSettleS := TIME_TO_REAL(tSettle) * 1.0E-3;          // 毫秒 → 秒（本行换算单位为 s）
ELSE
    tMove := DL_CALC_TIME_MAX;
    fSettleS := TIME_TO_REAL(DL_CALC_TIME_MAX) * 1.0E-3;
END_IF
tAccPhase    := T#0S;
tCruisePhase := T#0S;
tDecPhase    := T#0S;

// 段 2｜参数校验（非有限值先自比检测，再做域比较；公约 0.9）
bParamOk := (fDistance = fDistance) AND (fVelMax = fVelMax) AND (fAcc = fAcc)
            AND (fDec = fDec) AND (fVelStart = fVelStart)
            AND (ABS(fDistance) <= DL_CALC_INF_MAX) AND (ABS(fVelStart) <= DL_CALC_INF_MAX)
            AND (fVelMax > DL_CALC_VEL_FLOOR) AND (fVelMax <= DL_CALC_INF_MAX)
            AND (fAcc > DL_CALC_ACC_FLOOR) AND (fAcc <= DL_CALC_INF_MAX)
            AND (fDec > DL_CALC_ACC_FLOOR) AND (fDec <= DL_CALC_INF_MAX);
IF NOT bParamOk THEN
    FC_DL_CalcMoveTime := FALSE;                         // 参数非法：调用方必须先判返回值
    uErrorId           := 16#0004_0180;                  // 【信息级】参数非法
    tMove              := T#0S;
    RETURN;
END_IF

// 段 3｜输入归一化（负距离取绝对值，符号不影响耗时）
fDist    := ABS(fDistance);
fV0      := ABS(fVelStart);
fVmax    := fVelMax;
fA       := fAcc;
fDecUse  := fDec;

// 段 4｜距离为零：耗时即稳定延时
IF fDist <= DL_CALC_EPS THEN
    fVelPeak        := fV0;                              // 未移动，峰值速度即起始速度 [mm/s]
    bTriangular     := FALSE;                            // 总耗时保持默认值（= 稳定延时），无需重算
    uErrorId        := 16#0004_0182;                     // 【信息级】距离为零，耗时等于稳定延时
    RETURN;
END_IF

// 段 5｜起始速度已超上限：只能减速（接续定位的真实工况，不判失败）
IF fV0 > (fVmax + DL_CALC_EPS) THEN
    fDistStop := (fV0 * fV0) / (2.0 * fDecUse);           // 纯减速停车距离 [mm]，分母已验非零
    IF fDistStop >= (fDist - DL_CALC_EPS) THEN
        // 边减速边到点：到点速度为开方结果，被开方数防负数
        fRadicand := fV0 * fV0 - 2.0 * fDecUse * fDist;
        fRadicand := MAX(0.0, fRadicand);
        fVEnd     := SQRT(fRadicand);
        fTDec     := (fV0 - fVEnd) / fDecUse;             // 减速段耗时 [s]
        fTAcc     := 0.0;
        fTCruise  := 0.0;
    ELSE
        // 先减速到上限，再以匀速走完剩余行程
        fTDec      := (fV0 - fVmax) / fDecUse;            // 减速到上限耗时 [s]
        fDistDec   := (fV0 * fV0 - fVmax * fVmax) / (2.0 * fDecUse); // 减速段行程 [mm]
        fDistCruise:= fDist - fDistDec;
        IF fDistCruise < 0.0 THEN
            fDistCruise := 0.0;                           // 浮点残差钳零
        END_IF
        fTCruise   := fDistCruise / fVmax;                // 匀速段耗时 [s]，分母已验非零
        fTAcc      := 0.0;
        fDistAcc   := 0.0;
    END_IF
    fVelPeak := fV0;                                      // 峰值速度即起始速度 [mm/s]
    bTriangular := FALSE;
    uErrorId := 16#0004_0183;                             // 【信息级】起始速度超上限，按减速到点计算

ELSE
    // 段 6｜常规情形：先算临界距离，判梯形还是三角
    fDistCrit := (fVmax * fVmax - fV0 * fV0) / (2.0 * fA) + (fVmax * fVmax) / (2.0 * fDecUse);
    IF fDist >= (fDistCrit - DL_CALC_EPS) THEN
        // —— 梯形：可达速度上限 ——
        fTAcc      := (fVmax - fV0) / fA;                 // 加速段耗时 [s]
        fDistAcc   := (fVmax * fVmax - fV0 * fV0) / (2.0 * fA); // 加速段行程 [mm]
        fDistDec   := (fVmax * fVmax) / (2.0 * fDecUse);  // 减速段行程 [mm]
        fTDec      := fVmax / fDecUse;                    // 减速段耗时 [s]
        fDistCruise:= fDist - fDistAcc - fDistDec;
        IF fDistCruise < 0.0 THEN
            fDistCruise := 0.0;                           // 距离恰等于临界值的浮点残差：匀速段钳零
            uErrorId    := 16#0004_0181;                  // 【信息级】临界距离浮点残差，匀速段钳零
        END_IF
        fTCruise   := fDistCruise / fVmax;                // 匀速段耗时 [s]，分母已验非零
        fVelPeak   := fVmax;                              // 达到速度上限 [mm/s]
        bTriangular:= FALSE;
    ELSE
        // —— 三角：距离不足，峰速小于上限 ——
        fDenom    := fA + fDecUse;                        // 分母 > 0 已由校验保证
        fRadicand := 2.0 * fA * fDecUse * fDist + fDecUse * fV0 * fV0;
        fRadicand := MAX(0.0, fRadicand);
        fPeak     := SQRT(fRadicand / fDenom);            // 三角峰速 [mm/s]
        fVelPeak  := fPeak;
        fTAcc     := (fPeak - fV0) / fA;                  // 加速段耗时 [s]
        IF fTAcc < 0.0 THEN
            fTAcc := 0.0;                                 // 峰速低于起始速度时不加速（浮点残差防线）
        END_IF
        fTDec     := fPeak / fDecUse;                     // 减速段耗时 [s]
        fTCruise  := 0.0;                                 // 三角曲线无匀速段
        bTriangular := TRUE;                              // 三角退化：选型警示
        uErrorId  := 0;                                   // 正常三角退化不设码（属合法工况）
    END_IF
END_IF

// 段 7｜分段耗时换算（秒 → 毫秒，截断到毫秒，不做四舍五入以免累计偏大）
tAccPhase    := REAL_TO_TIME(fTAcc * DL_CALC_MS_SCALE);
tCruisePhase := REAL_TO_TIME(fTCruise * DL_CALC_MS_SCALE);
tDecPhase    := REAL_TO_TIME(fTDec * DL_CALC_MS_SCALE);

// 段 8｜总耗时合成与上限保护（防参数错填导致 HMI 时间控件溢出）
fTTotal := fTAcc + fTCruise + fTDec + fSettleS;
IF fTTotal > (TIME_TO_REAL(DL_CALC_TIME_MAX) * 1.0E-3) THEN
    tMove    := DL_CALC_TIME_MAX;                         // 超上限钳位
    uErrorId := 16#0004_0184;                             // 【信息级】结果超上限钳位
ELSE
    tMove := REAL_TO_TIME(fTTotal * DL_CALC_MS_SCALE);    // 总耗时 [ms]，含稳定延时
END_IF

// 段 9｜结果一致性复核（分段和不得超过总耗时，防浮点截断造成分段和大于总耗时）
IF (tAccPhase + tCruisePhase + tDecPhase) > tMove THEN
    tMove := tAccPhase + tCruisePhase + tDecPhase;        // 以分段和为准，保证上层相加自洽
END_IF

END_FUNCTION

(* ---- I_DL_MotionAxis.st ---- *)
(*==============================================================================
 * 组件名称 (Component)  : I_DL_MotionAxis
 * 所属子库 (Sublibrary) : DL_Motion
 * 当前版本 (Version)    : 1.0.0
 * 组件分类 (Category)   : 接口（INTERFACE）· 运动控制抽象契约 · Level 1 工艺层
 * 兼容性   (Platform)   : CODESYS 3.5 / TwinCAT 3 / 汇川 InoProShop / Schneider
 *                         Machine Expert；仅依赖 Standard.library，零厂商方言
 * 功能描述 (Function)   : 单轴运动控制标准抽象契约，按本库接口三段式公约
 *                         （0.11）组织：属性（PROPERTY GET）+ 方法（METHOD）
 *                         + 状态枚举。上层工艺块（点动器、工站、HMI 适配层）
 *                         仅依赖本接口引用，即可用同一套代码适配真实伺服
 *                         驱动、虚拟运动学仿真轴与第三方轴封装。
 * 方法数红线 (Budget)   : 方法共 6 个，恰在本库接口方法数红线（≤6）临界：
 *                         Enable / Reset / Stop / MoveAbsolute / MoveRelative /
 *                         MoveVelocity。回原（Homing）职责由后续轮次
 *                         FB_DL_AxisHomingSeq 承载，不入本接口。
 * 状态语义 (Semantics)  : E_DL_AxisState 按 PLCopen 轴状态模型 clean-room
 *                         重排：六态 + 禁用态，编号显式、间隔 10 预留扩展位
 *                         （R5 提取点 S-2④）。
 * 开源溯源 (Origin)     : plcopen / s7-motion。仅提取 PLCopen（TC5 接口规范
 *                         公开语义）轴状态名与命令动词、S7-1500 Motion Control
 *                         手册公开的工艺对象接口参数域；实现与命名 100% 自有，
 *                         clean-room，未参考任何厂商源码行。
 * 红线自检 (Redline)    : R1 ✓ 零全局变量表与外部变量引用 ｜ R2 ✓ 零物理地址直写
 *                         R3 ✓ 纯 IEC 61131-3 ｜ R4 N/A（契约件无运算）
 *                         R5 ✓ 全枚举项/方法参数双语注释 ｜ R6 N/A（接口无状态机）
 *                         R7 N/A（无实例调用）｜ R18 ✓ INTERFACE/END_INTERFACE 成对
 * 修订历史 (Revision)   :
 *   2026-11-15  v1.0.0  首版入库（Round 05 · DL_Motion 开库 · 接口契约件）
 *============================================================================*)

(*-----------------------------------------------------------------------------
 * 调用示例 (Instance guide)：
 *   VAR fbAxis : FB_DL_SingleAxis; END_VAR
 *   fbAxis();                                    // 先注入实参再周期调用
 *   bOk := fbAxis.Enable(bOn := TRUE);           // 上使能（MC_Power 语义）
 *   bOk := fbAxis.MoveAbsolute(fPos := 120.0, fVel := 50.0, fAcc := 500.0);
 *   fbAxis();                                    // 每周期调用驱动状态机
 *   IF fbAxis.bError THEN bOk2 := fbAxis.Reset(); END_IF
 *   上层注入：JogController.iAxis := fbAxis;（接口引用指向实现块实例）
 *   注意：方法全部非阻塞，仅置内部请求标志；跨周期动作由 FB 主体状态机执行。
 *----------------------------------------------------------------------------*)

(*-----------------------------------------------------------------------------
 * 常见误用与现场提示 (Field notes)：
 *   1 eState = eStopping 时一切运动指令被拒绝（MC_Stop 语义），上层不要
 *     在停止未完成前抢发定位指令，指令会直接返回 FALSE 而不排队。
 *   2 MoveRelative 的 fDist 带符号，负值即负向；MoveVelocity 的 fVel 同理，
 *     上层不必先换算方向再调用。
 *   3 bError 为派生式（仅反映 eErrorStop 态），信息级事件码只进 uErrorId，
 *     上层 HMI 报警分组时应同时读两者。
 *   4 bHomed 在本库当前版本恒为 FALSE 占位，回原由后续轮次组件驱动后置位；
 *     依赖回原联锁的工站请先行用安全限位方案替代。
 *   5 接口方法在实现块内必须逐个落地，任何新增实现块（真实驱动适配层）
 *     不得增删方法签名，否则破坏依赖本接口的全部上层块。
 *----------------------------------------------------------------------------*)

(*-----------------------------------------------------------------------------
 * 状态跃迁契约 (Transition contract)：
 *   实现块必须保证以下跃迁语义，供上层联锁与 HMI 依赖（本接口只定契约，
 *   实现块 FB_DL_SingleAxis 为参考实现，后续真实驱动适配层须逐条对齐）：
 *   1 eDisabled：唯一入态；仅 Enable(bOn=TRUE) 且驱动就绪可迁出至
 *     eStandstill，迁移后 bEnabled 必须为 TRUE。
 *   2 eStandstill：唯一可接收三种 Move 指令的稳态（速度模式可在
 *     eContinuousMotion 中改速）；下使能指令必须回到 eDisabled。
 *   3 eDiscreteMotion / eContinuousMotion：执行中收到 Stop 必须转入
 *     eStopping 受控减速，禁止直接跳变；到位/限位停车后回 eStandstill。
 *   4 eStopping：拒绝一切运动指令；停稳后回 eStandstill，期间不得有
 *     任何速度输出残留。
 *   5 eErrorStop：故障唯一锁存态，仅 Reset 且故障源消除后可退回
 *     eStandstill 或 eDisabled；bError 派生式仅反映本态。
 *   6 eHoming：预留态，回原序列由后续轮次 FB_DL_AxisHomingSeq 承载，
 *     实现块在本态内不得自行产生运动输出。
 *   7 任何跃迁语义变化视为 MAJOR 变更（见子库版本号约定），必须回写
 *     VERSION.md 迁移指引并同步依赖本接口的全部上层块。
 *   8 实现块文件头必须标注本接口版本依赖关系，接口升版时实现块同步
 *     升版并重跑验收向量基线（见前节）。
 *----------------------------------------------------------------------------*)

(*-----------------------------------------------------------------------------
 * 方法前置条件与返回值语义 (Method contract)：
 *   Enable(bOn) : BOOL    — 故障态或驱动未就绪时上使能请求返回 FALSE；
 *                           下使能请求恒受理（返回 TRUE），电平语义。
 *   Reset()     : BOOL    — 仅 eErrorStop 态受理返回 TRUE，其余态返回
 *                           FALSE；复位语义为"确认报警"，故障源未消除时
 *                           实现块不得真正退态。
 *   Stop()              — 受理后进入 eStopping；eErrorStop 态调用无效；
 *                           MC_Stop 语义：停止完成后仍拒绝新任务直至新
 *                           运动指令被显式受理。
 *   MoveAbsolute(fPos, fVel, fAcc) : BOOL
 *                         — 仅 eStandstill 受理；参数非法（非有限值、非
 *                           正值）或目标位超软限位返回 FALSE 且轴状态
 *                           不得发生任何改变。
 *   MoveRelative(fDist, fVel, fAcc) : BOOL
 *                         — 同上；fDist 带符号，目标落点 = 当前位置 +
 *                           fDist，落点越限即拒绝。
 *   MoveVelocity(fVel, fAcc) : BOOL
 *                         — eStandstill / eContinuousMotion 两态受理；
 *                           fVel 带符号，连续运动中再次调用为改速而非
 *                           重启。
 *----------------------------------------------------------------------------*)

(*-----------------------------------------------------------------------------
 * 实现块落地契约清单 (Implementer checklist)：
 *   后续任何新增实现块（真实伺服适配层、仿真轴、第三方轴包装类）实现
 *   本接口时必须逐条满足，否则视为违反库架构公约：
 *   1 七个 PROPERTY GET 必须全部落地，返回值与内部状态实时一致；
 *   2 六个 METHOD 必须全部落地且签名逐字一致，不得增删参数；
 *   3 方法内不得阻塞、不得跨扫描周期驻留临时状态，跨周期动作一律
 *     经内部请求标志由 FB 主体状态机执行；
 *   4 bError 必须为派生式且仅反映 eErrorStop 态，信息级事件只进
 *     uErrorId（R19/R21 公约）；
 *   5 实现块不得出现任何全局变量引用、外部变量声明或物理地址直写
 *     （R1/R2 红线），硬件差异全部由上层适配层吸收；
 *   6 状态枚举 E_DL_AxisState 的取值与语义不得重定义或扩展；
 *   7 故障码沿用 DL_Motion 族段位 16#0004_xxxx（信息级 01xx / 故障级
 *     02xx 起），不得自造码段。
 *----------------------------------------------------------------------------*)

(*-----------------------------------------------------------------------------
 * 验收向量基线 (Acceptance baseline)：
 *   本接口为契约件，验收向量在实现块上执行；实现块验收必须覆盖：
 *   1 正常跃迁链：Enable → eStandstill → MoveAbsolute → 到位回待机；
 *   2 非法状态兜底：内部状态被破坏后实现块 CASE+ELSE 兜底进 eErrorStop；
 *   3 运行中途插入跟踪脉冲：运动态插入 bTrack → 位置重同步 + 受控停车
 *     （R5 公约 0.1 必测向量）；
 *   4 指令门禁：eStopping/eErrorStop 态全部 Move 方法返回 FALSE 且
 *     轴状态不变；
 *   5 参数防御：非有限值与非正值参数被拒绝，接口引用未注入时上层
 *     调用不产生任何轴动作。
 *   6 一致性回归：实现块更新后须重跑 1~5 向量，任何跃迁语义变化视为
 *     MAJOR 变更（见子库版本号约定），必须回写 VERSION.md 迁移指引。
 *----------------------------------------------------------------------------*)

(*-----------------------------------------------------------------------------
 * 归属声明 (Ownership note)：
 *   E_DL_AxisState 为本接口契约的组成枚举，随本接口同文件发布（规格书
 *   第 6 节交付约定：接口与其枚举同文件，头注释注明归属）。导入 .st 后
 *   枚举全局可见，实现块 FB_DL_SingleAxis 与上层工艺块直接引用。
 *----------------------------------------------------------------------------*)

{attribute 'strict'}
{attribute 'qualified_only'}
TYPE E_DL_AxisState :
(
    eDisabled         := 0,    // 禁用：伺服未上使能，输出级切断 / Disabled: servo not enabled, outputs cut off
    eStandstill       := 10,   // 待机：已使能且静止就绪，可接收运动指令 / Standstill: enabled and stationary, ready for motion commands
    eHoming           := 20,   // 回原中：回原点序列执行中（后续轮次组件承载） / Homing: homing sequence in progress (reserved)
    eDiscreteMotion   := 30,   // 离散运动中：绝对/相对定位执行中 / Discrete motion: absolute or relative positioning active
    eContinuousMotion := 40,   // 连续运动中：速度模式执行中 / Continuous motion: velocity mode active
    eStopping         := 50,   // 受控停止中：按减速度斜坡停车，拒绝新任务 / Stopping: controlled deceleration, new tasks rejected
    eErrorStop        := 60    // 故障停机：报警锁存，仅 Reset 可退回 / Error stop: fault latched, only Reset can leave
) UINT;
END_TYPE

INTERFACE I_DL_MotionAxis

(* —— 段 1｜属性（PROPERTY GET）：状态只读出口，实现块一一落地 —— *)
PROPERTY eState    : E_DL_AxisState   // 当前轴状态（Current axis state），枚举见 E_DL_AxisState
END_PROPERTY
PROPERTY fPosition : REAL             // 当前位置（Current position）[mm 或 deg，单位由实现组态注释约定]
END_PROPERTY
PROPERTY fVelocity : REAL             // 当前速度（Current velocity）[mm/s 或 deg/s]，带符号，负值=负向
END_PROPERTY
PROPERTY bEnabled  : BOOL             // 使能状态（Enabled status），TRUE=伺服已上使能
END_PROPERTY
PROPERTY bHomed    : BOOL             // 回原完成（Homed status），TRUE=坐标系已建立
END_PROPERTY
PROPERTY bError    : BOOL             // 故障锁存（Error latched），TRUE=处于 eErrorStop 态
END_PROPERTY
PROPERTY uErrorId  : UDINT            // 末次事件码（Last error code），信息级码不置 bError
END_PROPERTY

(* —— 段 2｜方法（METHOD）：命令入口，全部非阻塞单发化 —— *)
METHOD Enable : BOOL                       // 使能请求（Enable request），MC_Power 语义
VAR_INPUT
    bOn : BOOL;                            // 使能电平（Enable on/off），TRUE=上使能请求 / FALSE=下使能请求
END_VAR

    END_METHOD

METHOD Reset : BOOL                        // 故障复位（Fault reset），MC_Reset 语义，确认报警
VAR_INPUT
END_VAR

    END_METHOD

METHOD Stop                                // 受控停止（Controlled stop），MC_Stop 语义：停车并拒绝新任务
VAR_INPUT
END_VAR

    END_METHOD

METHOD MoveAbsolute : BOOL                 // 绝对定位（Move absolute）
VAR_INPUT
    fPos : REAL;                           // 目标绝对位置（Target absolute position）[mm 或 deg]
    fVel : REAL;                           // 运行速度（Run velocity）[mm/s]，正值，超上限自动钳位
    fAcc : REAL;                           // 加/减速度（Acceleration and deceleration）[mm/s²]，正值
END_VAR

    END_METHOD

METHOD MoveRelative : BOOL                 // 相对定位（Move relative）
VAR_INPUT
    fDist : REAL;                          // 相对位移（Relative distance）[mm]，带符号，负值=负向
    fVel  : REAL;                          // 运行速度（Run velocity）[mm/s]，正值
    fAcc  : REAL;                          // 加/减速度（Acceleration and deceleration）[mm/s²]，正值
END_VAR

    END_METHOD

METHOD MoveVelocity : BOOL                 // 速度模式（Move velocity），可在连续运动中改速
VAR_INPUT
    fVel : REAL;                           // 目标速度（Target velocity）[mm/s]，带符号，负值=负向
    fAcc : REAL;                           // 加/减速度（Acceleration and deceleration）[mm/s²]，正值
END_VAR

    END_METHOD
END_INTERFACE
